(* IEC 61131-3 sources: plc-st-coding-agent/progress/evidence/f14_v10_full_20261113/jobs/codex_minimax-m27 (part 6) *)

(* ---- public-medium-08.raw_candidate_04.st ---- *)
(* ENGINEERING_CONTRACT
   PUB001: Parse dotted-decimal IPv4, validate 4 numeric segments 0-255
   PUB002: Network byte order assembly (MSB=first segment)
   PUB003: Invalid input → ipValue=0 (malformed, nondigit, wrong count, OOR)
   PUB004: Valid 0.0.0.0 also produces 0 (by assembly)

   State retention: None (stateless function block)
   Reset behavior: None (no reset input specified)
   First scan: Same as subsequent (no edge memory)

   Bug fix: Reject empty segments (consecutive delimiters like "1..2.3")
   by tracking nonempty digit accumulation per segment
*)

(* CONTRACT_RULES [] *)

FUNCTION_BLOCK IPv4_Parse
VAR_INPUT
    ipText : STRING(254);
END_VAR
VAR_OUTPUT
    ipValue : UDINT := 0;
END_VAR
VAR
    tmp_pos : UDINT;
    tmp_seg_idx : UDINT;
    tmp_char : BYTE;
    tmp_seg_val : UDINT;
    tmp_result : UDINT;
    tmp_seg_nonempty : BOOL;
END_VAR

tmp_pos := 0;
tmp_seg_idx := 0;
tmp_result := 0;
tmp_seg_val := 0;
tmp_seg_nonempty := FALSE;

WHILE tmp_pos < LEN(ipText) DO
    tmp_char := ipText[tmp_pos];

    IF tmp_char >= 48 AND tmp_char <= 57 THEN
        tmp_seg_val := tmp_seg_val * 10 + TO_UDINT(tmp_char - 48);

        IF tmp_seg_val > 255 THEN
            ipValue := 0;
            RETURN;
        END_IF;

        tmp_seg_nonempty := TRUE;
        tmp_pos := tmp_pos + 1;

    ELSIF tmp_char = 46 THEN

        IF NOT tmp_seg_nonempty THEN
            ipValue := 0;
            RETURN;
        END_IF;

        IF tmp_seg_idx >= 3 THEN
            ipValue := 0;
            RETURN;
        END_IF;

        CASE tmp_seg_idx OF
            0: tmp_result := SHL(tmp_seg_val, 24);
            1: tmp_result := tmp_result OR SHL(tmp_seg_val, 16);
            2: tmp_result := tmp_result OR SHL(tmp_seg_val, 8);
        END_CASE;

        tmp_seg_idx := tmp_seg_idx + 1;
        tmp_seg_val := 0;
        tmp_seg_nonempty := FALSE;
        tmp_pos := tmp_pos + 1;
    ELSE

        ipValue := 0;
        RETURN;
    END_IF;
END_WHILE;

IF tmp_seg_idx <> 3 THEN
    ipValue := 0;
ELSE
    tmp_result := tmp_result OR tmp_seg_val;
    ipValue := tmp_result;
END_IF;

END_FUNCTION_BLOCK

(* ---- self-easy-01.candidate_01.st ---- *)
(*
ENGINEERING_CONTRACT
================================================================
Output: avgOut (REAL)
─────────────────────────────────────────────────────────────────
Activation:    Computed every scan when enable AND avgEnable AND count > 0
Retention:     Held when enable=FALSE, avgEnable=FALSE, or count<=0
Reset:         No explicit reset; cold-start avgOut initializes to 0.0
Same-scan:     All inputs evaluated together; final timer state used
Units/bounds:  count: 0..8 clamped to 1..8 for division, sum: DINT
─────────────────────────────────────────────────────────────────
PUB001: enable=TRUE updates avgOut; enable=FALSE retains prev
PUB002: avgEnable input
PUB003: values array[1..8] of INT, 1-indexed sample storage
PUB004: count input INT
PUB005: avgOut output REAL, no rounding to integer
PUB006: count=0 -> no division by zero, avgOut unchanged
PUB007: count>8 -> use only first 8 samples, no out-of-bounds
PUB008: avgEnable=FALSE -> avgOut unchanged (retain)
PUB009: DINT/LINT summation to prevent INT overflow
PUB010: REAL output preserves original precision
================================================================
*)

(* CONTRACT_RULES [] *)

FUNCTION_BLOCK FB
VAR_INPUT
    enable    : BOOL;
    values    : ARRAY[1..8] OF INT;
    count     : INT;
    avgEnable : BOOL;
END_VAR
VAR_OUTPUT
    avgOut    : REAL := 0.0;
END_VAR
VAR
    tmp_sum   : DINT;
    tmp_count : INT;
END_VAR

tmp_count := count;
IF tmp_count < 1 THEN
    tmp_count := 0;
ELSIF tmp_count > 8 THEN
    tmp_count := 8;
END_IF;

IF enable AND avgEnable AND (tmp_count > 0) THEN
    tmp_sum := 0;
    IF tmp_count >= 1 THEN
        tmp_sum := tmp_sum + TO_DINT(values[1]);
    END_IF;
    IF tmp_count >= 2 THEN
        tmp_sum := tmp_sum + TO_DINT(values[2]);
    END_IF;
    IF tmp_count >= 3 THEN
        tmp_sum := tmp_sum + TO_DINT(values[3]);
    END_IF;
    IF tmp_count >= 4 THEN
        tmp_sum := tmp_sum + TO_DINT(values[4]);
    END_IF;
    IF tmp_count >= 5 THEN
        tmp_sum := tmp_sum + TO_DINT(values[5]);
    END_IF;
    IF tmp_count >= 6 THEN
        tmp_sum := tmp_sum + TO_DINT(values[6]);
    END_IF;
    IF tmp_count >= 7 THEN
        tmp_sum := tmp_sum + TO_DINT(values[7]);
    END_IF;
    IF tmp_count >= 8 THEN
        tmp_sum := tmp_sum + TO_DINT(values[8]);
    END_IF;
    avgOut := TO_REAL(tmp_sum) / TO_REAL(tmp_count);
END_IF;
END_FUNCTION_BLOCK

(* ---- self-easy-01.raw_candidate_01.st ---- *)
(*
ENGINEERING_CONTRACT
================================================================
Output: avgOut (REAL)
─────────────────────────────────────────────────────────────────
Activation:    Computed every scan when enable AND avgEnable AND count > 0
Retention:     Held when enable=FALSE, avgEnable=FALSE, or count<=0
Reset:         No explicit reset; cold-start avgOut initializes to 0.0
Same-scan:     All inputs evaluated together; final timer state used
Units/bounds:  count: 0..8 clamped to 1..8 for division, sum: DINT
─────────────────────────────────────────────────────────────────
PUB001: enable=TRUE updates avgOut; enable=FALSE retains prev
PUB002: avgEnable input
PUB003: values array[1..8] of INT, 1-indexed sample storage
PUB004: count input INT
PUB005: avgOut output REAL, no rounding to integer
PUB006: count=0 -> no division by zero, avgOut unchanged
PUB007: count>8 -> use only first 8 samples, no out-of-bounds
PUB008: avgEnable=FALSE -> avgOut unchanged (retain)
PUB009: DINT/LINT summation to prevent INT overflow
PUB010: REAL output preserves original precision
================================================================
*)

(* CONTRACT_RULES [] *)

FUNCTION_BLOCK FB
VAR_INPUT
    enable    : BOOL;
    values    : ARRAY[1..8] OF INT;
    count     : INT;
    avgEnable : BOOL;
END_VAR
VAR_OUTPUT
    avgOut    : REAL := 0.0;
END_VAR
VAR
    tmp_sum   : DINT;
    tmp_count : INT;
END_VAR

tmp_count := count;
IF tmp_count < 1 THEN
    tmp_count := 0;
ELSIF tmp_count > 8 THEN
    tmp_count := 8;
END_IF;

IF enable AND avgEnable AND (tmp_count > 0) THEN
    tmp_sum := 0;
    IF tmp_count >= 1 THEN
        tmp_sum := tmp_sum + TO_DINT(values[1]);
    END_IF;
    IF tmp_count >= 2 THEN
        tmp_sum := tmp_sum + TO_DINT(values[2]);
    END_IF;
    IF tmp_count >= 3 THEN
        tmp_sum := tmp_sum + TO_DINT(values[3]);
    END_IF;
    IF tmp_count >= 4 THEN
        tmp_sum := tmp_sum + TO_DINT(values[4]);
    END_IF;
    IF tmp_count >= 5 THEN
        tmp_sum := tmp_sum + TO_DINT(values[5]);
    END_IF;
    IF tmp_count >= 6 THEN
        tmp_sum := tmp_sum + TO_DINT(values[6]);
    END_IF;
    IF tmp_count >= 7 THEN
        tmp_sum := tmp_sum + TO_DINT(values[7]);
    END_IF;
    IF tmp_count >= 8 THEN
        tmp_sum := tmp_sum + TO_DINT(values[8]);
    END_IF;
    avgOut := TO_REAL(tmp_sum) / TO_REAL(tmp_count);
END_IF;
END_FUNCTION_BLOCK

(* ---- self-easy-02.candidate_01.st ---- *)
FUNCTION_BLOCK FB
VAR_INPUT
    tankLevel   : REAL;
    outletFlow  : REAL;
    inletPermit : BOOL;
    resetBtn    : BOOL;
END_VAR
VAR_OUTPUT
    pumpRun        : BOOL;
    alarmHigh      : BOOL;
    alarmLow       : BOOL;
    outletValveOpen: BOOL;
END_VAR
VAR
    prevResetBtn   : BOOL := FALSE;
    prevAlarmHigh  : BOOL := FALSE;
    prevAlarmLow   : BOOL := FALSE;
    firstScan      : BOOL := TRUE;
END_VAR
(* ENGINEERING_CONTRACT
 * ┌──────────────────┬─────────────────────────────────────────────────────────┐
 * │ alarmHigh        │ SET: tankLevel >= 85.0 (same scan priority)             │
 * │                  │ HOLD: until resetBtn rising edge AND tankLevel < 85.0   │
 * │                  │ RESET: only when safe condition cleared first           │
 * │                  │ UNITS: dimensionless % [0..100]                         │
 * ├──────────────────┼─────────────────────────────────────────────────────────┤
 * │ alarmLow         │ SET: tankLevel <= 15.0 (same scan priority)             │
 * │                  │ HOLD: until resetBtn rising edge AND tankLevel > 15.0   │
 * │                  │ RESET: only when safe condition cleared first           │
 * │                  │ UNITS: dimensionless % [0..100]                         │
 * ├──────────────────┼─────────────────────────────────────────────────────────┤
 * │ pumpRun          │ ACTIVATION: inletPermit=TRUE AND alarmHigh=FALSE AND alarmLow=FALSE │
 * │                  │ DEACTIVATION: any alarm active OR inletPermit=FALSE     │
 * │                  │ PRIORITY: stop-before-start, same-scan final state      │
 * │                  │ UNITS: command signal (BOOL)                            │
 * ├──────────────────┼─────────────────────────────────────────────────────────┤
 * │ outletValveOpen  │ ACTIVATION: alarmLow=FALSE (normal + alarmHigh-only)    │
 * │                  │ DEACTIVATION: alarmLow=TRUE                             │
 * │                  │ PRIORITY: latch follows alarmLow, no reset edge effect  │
 * │                  │ UNITS: command signal (BOOL)                            │
 * ├──────────────────┼─────────────────────────────────────────────────────────┤
 * │ resetBtn edge    │ DETECT: rising(TRUE), firstScan treated as FALSE->FALSE  │
 * │                  │ RETENTION: holding across level change does NOT trigger │
 * │                  │ UNITS: edge-detected per scan                           │
 * └──────────────────┴─────────────────────────────────────────────────────────┘
 * PUB refs: 85%/15% thresholds PUB003, latch PUB004, reset edge PUB005,
 *           pump interlock PUB006, valve PUB007, inlet permit PUB008
 *)
BEGIN
    (* Detect rising edge on resetBtn; first scan treats btn as FALSE *)
    IF firstScan THEN
        firstScan := FALSE;
    END_IF;

    (* Step 1: Update alarmHigh - immediate latch on danger condition *)
    IF tankLevel >= 85.0 THEN
        alarmHigh := TRUE;
    ELSIF resetBtn AND NOT prevResetBtn AND tankLevel < 85.0 THEN
        alarmHigh := FALSE;
    END_IF;

    (* Step 2: Update alarmLow - immediate latch on danger condition *)
    IF tankLevel <= 15.0 THEN
        alarmLow := TRUE;
    ELSIF resetBtn AND NOT prevResetBtn AND tankLevel > 15.0 THEN
        alarmLow := FALSE;
    END_IF;

    (* Step 3: pumpRun - stop before start, all conditions same scan *)
    IF alarmHigh OR alarmLow OR NOT inletPermit THEN
        pumpRun := FALSE;
    ELSE
        pumpRun := TRUE;
    END_IF;

    (* Step 4: outletValveOpen - inverse of alarmLow *)
    outletValveOpen := NOT alarmLow;

    (* Step 5: Store previous states for next scan edge detection *)
    prevResetBtn  := resetBtn;
    prevAlarmHigh := alarmHigh;
    prevAlarmLow  := alarmLow;
END_FUNCTION_BLOCK

(* ---- self-easy-02.candidate_02.st ---- *)
FUNCTION_BLOCK FB
VAR_INPUT
    tankLevel   : REAL;
    outletFlow  : REAL;
    inletPermit : BOOL;
    resetBtn    : BOOL;
END_VAR
VAR_OUTPUT
    pumpRun        : BOOL;
    alarmHigh      : BOOL;
    alarmLow       : BOOL;
    outletValveOpen: BOOL;
END_VAR
VAR
    prevResetBtn   : BOOL := FALSE;
    prevAlarmHigh  : BOOL := FALSE;
    prevAlarmLow   : BOOL := FALSE;
    firstScan      : BOOL := TRUE;
END_VAR
(* ENGINEERING_CONTRACT
 * ┌──────────────────┬─────────────────────────────────────────────────────────┐
 * │ alarmHigh        │ SET: tankLevel >= 85.0 (same scan priority)             │
 * │                  │ HOLD: until resetBtn rising edge AND tankLevel < 85.0   │
 * │                  │ RESET: only when safe condition cleared first           │
 * │                  │ UNITS: dimensionless % [0..100]                         │
 * ├──────────────────┼─────────────────────────────────────────────────────────┤
 * │ alarmLow         │ SET: tankLevel <= 15.0 (same scan priority)             │
 * │                  │ HOLD: until resetBtn rising edge AND tankLevel > 15.0   │
 * │                  │ RESET: only when safe condition cleared first           │
 * │                  │ UNITS: dimensionless % [0..100]                         │
 * ├──────────────────┼─────────────────────────────────────────────────────────┤
 * │ pumpRun          │ ACTIVATION: inletPermit=TRUE AND alarmHigh=FALSE AND alarmLow=FALSE │
 * │                  │ DEACTIVATION: any alarm active OR inletPermit=FALSE     │
 * │                  │ PRIORITY: stop-before-start, same-scan final state      │
 * │                  │ UNITS: command signal (BOOL)                            │
 * ├──────────────────┼─────────────────────────────────────────────────────────┤
 * │ outletValveOpen  │ ACTIVATION: alarmLow=FALSE (normal + alarmHigh-only)    │
 * │                  │ DEACTIVATION: alarmLow=TRUE                             │
 * │                  │ PRIORITY: latch follows alarmLow, no reset edge effect  │
 * │                  │ UNITS: command signal (BOOL)                            │
 * ├──────────────────┼─────────────────────────────────────────────────────────┤
 * │ resetBtn edge    │ DETECT: rising(TRUE), firstScan treated as FALSE->FALSE  │
 * │                  │ RETENTION: holding across level change does NOT trigger │
 * │                  │ UNITS: edge-detected per scan                           │
 * └──────────────────┴─────────────────────────────────────────────────────────┘
 * PUB refs: 85%/15% thresholds PUB003, latch PUB004, reset edge PUB005,
 *           pump interlock PUB006, valve PUB007, inlet permit PUB008
 *)
BEGIN
    (* Step 1: Update alarmHigh - immediate latch on danger condition *)
    IF tankLevel >= 85.0 THEN
        alarmHigh := TRUE;
    ELSIF resetBtn AND NOT prevResetBtn AND NOT firstScan AND tankLevel < 85.0 THEN
        alarmHigh := FALSE;
    END_IF;

    (* Step 2: Update alarmLow - immediate latch on danger condition *)
    IF tankLevel <= 15.0 THEN
        alarmLow := TRUE;
    ELSIF resetBtn AND NOT prevResetBtn AND NOT firstScan AND tankLevel > 15.0 THEN
        alarmLow := FALSE;
    END_IF;

    (* Step 3: pumpRun - stop before start, all conditions same scan *)
    IF alarmHigh OR alarmLow OR NOT inletPermit THEN
        pumpRun := FALSE;
    ELSE
        pumpRun := TRUE;
    END_IF;

    (* Step 4: outletValveOpen - inverse of alarmLow *)
    outletValveOpen := NOT alarmLow;

    (* Step 5: Store previous states for next scan *)
    prevResetBtn  := resetBtn;
    prevAlarmHigh := alarmHigh;
    prevAlarmLow  := alarmLow;
    firstScan     := FALSE;
END_FUNCTION_BLOCK

(* ---- self-easy-02.candidate_03.st ---- *)
FUNCTION_BLOCK FB
VAR_INPUT
    tankLevel   : REAL;
    outletFlow  : REAL;
    inletPermit : BOOL;
    resetBtn    : BOOL;
END_VAR
VAR_OUTPUT
    pumpRun        : BOOL;
    alarmHigh      : BOOL;
    alarmLow       : BOOL;
    outletValveOpen: BOOL;
END_VAR
VAR
    prevResetBtn : BOOL := FALSE;
END_VAR
(* ENGINEERING_CONTRACT *)
(* alarmHigh: SET at tankLevel>=85.0 (same-scan priority). HOLD until resetBtn rising AND tankLevel<85.0. RESET only when safe first. *)
(* alarmLow:  SET at tankLevel<=15.0 (same-scan priority). HOLD until resetBtn rising AND tankLevel>15.0. RESET only when safe first. *)
(* pumpRun:   ACT when inletPermit=TRUE AND alarmHigh=FALSE AND alarmLow=FALSE. STOP on any alarm or !inletPermit. *)
(* outletValveOpen: ON when alarmLow=FALSE. OFF when alarmLow=TRUE. No reset edge effect. *)
(* resetBtn:  Rising edge detection, firstScan=FALSE. Holding across level change does NOT re-trigger. *)
BEGIN
    (* Update alarmHigh *)
    IF tankLevel >= 85.0 THEN
        alarmHigh := TRUE;
    ELSIF resetBtn AND NOT prevResetBtn AND tankLevel < 85.0 THEN
        alarmHigh := FALSE;
    END_IF;

    (* Update alarmLow *)
    IF tankLevel <= 15.0 THEN
        alarmLow := TRUE;
    ELSIF resetBtn AND NOT prevResetBtn AND tankLevel > 15.0 THEN
        alarmLow := FALSE;
    END_IF;

    (* pumpRun: stop before start *)
    IF alarmHigh OR alarmLow OR NOT inletPermit THEN
        pumpRun := FALSE;
    ELSE
        pumpRun := TRUE;
    END_IF;

    (* outletValveOpen: inverse of alarmLow *)
    outletValveOpen := NOT alarmLow;

    (* Store previous state *)
    prevResetBtn := resetBtn;
END_FUNCTION_BLOCK
(* CONTRACT_RULES [] *)

(* ---- self-easy-02.candidate_04.st ---- *)
FUNCTION_BLOCK FB
VAR_INPUT
    tankLevel   : REAL;
    outletFlow  : REAL;
    inletPermit : BOOL;
    resetBtn    : BOOL;
END_VAR
VAR_OUTPUT
    pumpRun        : BOOL;
    alarmHigh      : BOOL;
    alarmLow       : BOOL;
    outletValveOpen: BOOL;
END_VAR
VAR
    prevResetBtn   : BOOL := FALSE;
    firstScan      : BOOL := TRUE;
END_VAR
(* ENGINEERING_CONTRACT
 * ┌──────────────────┬─────────────────────────────────────────────────────────┐
 * │ alarmHigh        │ SET: tankLevel >= 85.0 (same scan priority)             │
 * │                  │ HOLD: until resetBtn rising edge AND tankLevel < 85.0   │
 * │                  │ RESET: only when safe condition cleared first           │
 * │                  │ UNITS: dimensionless % [0..100]                         │
 * ├──────────────────┼─────────────────────────────────────────────────────────┤
 * │ alarmLow         │ SET: tankLevel <= 15.0 (same scan priority)             │
 * │                  │ HOLD: until resetBtn rising edge AND tankLevel > 15.0   │
 * │                  │ RESET: only when safe condition cleared first           │
 * │                  │ UNITS: dimensionless % [0..100]                         │
 * ├──────────────────┼─────────────────────────────────────────────────────────┤
 * │ pumpRun          │ ACTIVATION: inletPermit=TRUE AND alarmHigh=FALSE AND alarmLow=FALSE │
 * │                  │ DEACTIVATION: any alarm active OR inletPermit=FALSE     │
 * │                  │ PRIORITY: stop-before-start, same-scan final state      │
 * │                  │ UNITS: command signal (BOOL)                            │
 * ├──────────────────┼─────────────────────────────────────────────────────────┤
 * │ outletValveOpen  │ ACTIVATION: alarmLow=FALSE (normal + alarmHigh-only)    │
 * │                  │ DEACTIVATION: alarmLow=TRUE                             │
 * │                  │ PRIORITY: latch follows alarmLow, no reset edge effect  │
 * │                  │ UNITS: command signal (BOOL)                            │
 * ├──────────────────┼─────────────────────────────────────────────────────────┤
 * │ resetBtn edge    │ DETECT: rising(TRUE), firstScan treated as FALSE->FALSE  │
 * │                  │ RETENTION: holding across level change does NOT trigger │
 * │                  │ UNITS: edge-detected per scan                           │
 * └──────────────────┴─────────────────────────────────────────────────────────┘
 * PUB refs: 85%/15% thresholds PUB003, latch PUB004, reset edge PUB005,
 *           pump interlock PUB006, valve PUB007, inlet permit PUB008
 *)
BEGIN
    IF firstScan THEN
        firstScan := FALSE;
        prevResetBtn := FALSE;
    END_IF;

    IF tankLevel >= 85.0 THEN
        alarmHigh := TRUE;
    ELSIF resetBtn AND NOT prevResetBtn AND tankLevel < 85.0 THEN
        alarmHigh := FALSE;
    END_IF;

    IF tankLevel <= 15.0 THEN
        alarmLow := TRUE;
    ELSIF resetBtn AND NOT prevResetBtn AND tankLevel > 15.0 THEN
        alarmLow := FALSE;
    END_IF;

    IF alarmHigh OR alarmLow OR NOT inletPermit THEN
        pumpRun := FALSE;
    ELSE
        pumpRun := TRUE;
    END_IF;

    outletValveOpen := NOT alarmLow;

    prevResetBtn := resetBtn;
END_FUNCTION_BLOCK
(* CONTRACT_RULES [] *)

(* ---- self-easy-02.raw_candidate_01.st ---- *)
FUNCTION_BLOCK FB
VAR_INPUT
    tankLevel   : REAL;
    outletFlow  : REAL;
    inletPermit : BOOL;
    resetBtn    : BOOL;
END_VAR
VAR_OUTPUT
    pumpRun        : BOOL;
    alarmHigh      : BOOL;
    alarmLow       : BOOL;
    outletValveOpen: BOOL;
END_VAR
VAR
    prevResetBtn   : BOOL := FALSE;
    prevAlarmHigh  : BOOL := FALSE;
    prevAlarmLow   : BOOL := FALSE;
    firstScan      : BOOL := TRUE;
END_VAR
(* ENGINEERING_CONTRACT
 * ┌──────────────────┬─────────────────────────────────────────────────────────┐
 * │ alarmHigh        │ SET: tankLevel >= 85.0 (same scan priority)             │
 * │                  │ HOLD: until resetBtn rising edge AND tankLevel < 85.0   │
 * │                  │ RESET: only when safe condition cleared first           │
 * │                  │ UNITS: dimensionless % [0..100]                         │
 * ├──────────────────┼─────────────────────────────────────────────────────────┤
 * │ alarmLow         │ SET: tankLevel <= 15.0 (same scan priority)             │
 * │                  │ HOLD: until resetBtn rising edge AND tankLevel > 15.0   │
 * │                  │ RESET: only when safe condition cleared first           │
 * │                  │ UNITS: dimensionless % [0..100]                         │
 * ├──────────────────┼─────────────────────────────────────────────────────────┤
 * │ pumpRun          │ ACTIVATION: inletPermit=TRUE AND alarmHigh=FALSE AND alarmLow=FALSE │
 * │                  │ DEACTIVATION: any alarm active OR inletPermit=FALSE     │
 * │                  │ PRIORITY: stop-before-start, same-scan final state      │
 * │                  │ UNITS: command signal (BOOL)                            │
 * ├──────────────────┼─────────────────────────────────────────────────────────┤
 * │ outletValveOpen  │ ACTIVATION: alarmLow=FALSE (normal + alarmHigh-only)    │
 * │                  │ DEACTIVATION: alarmLow=TRUE                             │
 * │                  │ PRIORITY: latch follows alarmLow, no reset edge effect  │
 * │                  │ UNITS: command signal (BOOL)                            │
 * ├──────────────────┼─────────────────────────────────────────────────────────┤
 * │ resetBtn edge    │ DETECT: rising(TRUE), firstScan treated as FALSE->FALSE  │
 * │                  │ RETENTION: holding across level change does NOT trigger │
 * │                  │ UNITS: edge-detected per scan                           │
 * └──────────────────┴─────────────────────────────────────────────────────────┘
 * PUB refs: 85%/15% thresholds PUB003, latch PUB004, reset edge PUB005,
 *           pump interlock PUB006, valve PUB007, inlet permit PUB008
 *)
BEGIN
    (* Detect rising edge on resetBtn; first scan treats btn as FALSE *)
    IF firstScan THEN
        firstScan := FALSE;
    END_IF;

    (* Step 1: Update alarmHigh - immediate latch on danger condition *)
    IF tankLevel >= 85.0 THEN
        alarmHigh := TRUE;
    ELSIF resetBtn AND NOT prevResetBtn AND tankLevel < 85.0 THEN
        alarmHigh := FALSE;
    END_IF;

    (* Step 2: Update alarmLow - immediate latch on danger condition *)
    IF tankLevel <= 15.0 THEN
        alarmLow := TRUE;
    ELSIF resetBtn AND NOT prevResetBtn AND tankLevel > 15.0 THEN
        alarmLow := FALSE;
    END_IF;

    (* Step 3: pumpRun - stop before start, all conditions same scan *)
    IF alarmHigh OR alarmLow OR NOT inletPermit THEN
        pumpRun := FALSE;
    ELSE
        pumpRun := TRUE;
    END_IF;

    (* Step 4: outletValveOpen - inverse of alarmLow *)
    outletValveOpen := NOT alarmLow;

    (* Step 5: Store previous states for next scan edge detection *)
    prevResetBtn  := resetBtn;
    prevAlarmHigh := alarmHigh;
    prevAlarmLow  := alarmLow;
END_FUNCTION_BLOCK

(* ---- self-easy-02.raw_candidate_02.st ---- *)
FUNCTION_BLOCK FB
VAR_INPUT
    tankLevel   : REAL;
    outletFlow  : REAL;
    inletPermit : BOOL;
    resetBtn    : BOOL;
END_VAR
VAR_OUTPUT
    pumpRun        : BOOL;
    alarmHigh      : BOOL;
    alarmLow       : BOOL;
    outletValveOpen: BOOL;
END_VAR
VAR
    prevResetBtn   : BOOL := FALSE;
    prevAlarmHigh  : BOOL := FALSE;
    prevAlarmLow   : BOOL := FALSE;
    firstScan      : BOOL := TRUE;
END_VAR
(* ENGINEERING_CONTRACT
 * ┌──────────────────┬─────────────────────────────────────────────────────────┐
 * │ alarmHigh        │ SET: tankLevel >= 85.0 (same scan priority)             │
 * │                  │ HOLD: until resetBtn rising edge AND tankLevel < 85.0   │
 * │                  │ RESET: only when safe condition cleared first           │
 * │                  │ UNITS: dimensionless % [0..100]                         │
 * ├──────────────────┼─────────────────────────────────────────────────────────┤
 * │ alarmLow         │ SET: tankLevel <= 15.0 (same scan priority)             │
 * │                  │ HOLD: until resetBtn rising edge AND tankLevel > 15.0   │
 * │                  │ RESET: only when safe condition cleared first           │
 * │                  │ UNITS: dimensionless % [0..100]                         │
 * ├──────────────────┼─────────────────────────────────────────────────────────┤
 * │ pumpRun          │ ACTIVATION: inletPermit=TRUE AND alarmHigh=FALSE AND alarmLow=FALSE │
 * │                  │ DEACTIVATION: any alarm active OR inletPermit=FALSE     │
 * │                  │ PRIORITY: stop-before-start, same-scan final state      │
 * │                  │ UNITS: command signal (BOOL)                            │
 * ├──────────────────┼─────────────────────────────────────────────────────────┤
 * │ outletValveOpen  │ ACTIVATION: alarmLow=FALSE (normal + alarmHigh-only)    │
 * │                  │ DEACTIVATION: alarmLow=TRUE                             │
 * │                  │ PRIORITY: latch follows alarmLow, no reset edge effect  │
 * │                  │ UNITS: command signal (BOOL)                            │
 * ├──────────────────┼─────────────────────────────────────────────────────────┤
 * │ resetBtn edge    │ DETECT: rising(TRUE), firstScan treated as FALSE->FALSE  │
 * │                  │ RETENTION: holding across level change does NOT trigger │
 * │                  │ UNITS: edge-detected per scan                           │
 * └──────────────────┴─────────────────────────────────────────────────────────┘
 * PUB refs: 85%/15% thresholds PUB003, latch PUB004, reset edge PUB005,
 *           pump interlock PUB006, valve PUB007, inlet permit PUB008
 *)
BEGIN
    (* Step 1: Update alarmHigh - immediate latch on danger condition *)
    IF tankLevel >= 85.0 THEN
        alarmHigh := TRUE;
    ELSIF resetBtn AND NOT prevResetBtn AND NOT firstScan AND tankLevel < 85.0 THEN
        alarmHigh := FALSE;
    END_IF;

    (* Step 2: Update alarmLow - immediate latch on danger condition *)
    IF tankLevel <= 15.0 THEN
        alarmLow := TRUE;
    ELSIF resetBtn AND NOT prevResetBtn AND NOT firstScan AND tankLevel > 15.0 THEN
        alarmLow := FALSE;
    END_IF;

    (* Step 3: pumpRun - stop before start, all conditions same scan *)
    IF alarmHigh OR alarmLow OR NOT inletPermit THEN
        pumpRun := FALSE;
    ELSE
        pumpRun := TRUE;
    END_IF;

    (* Step 4: outletValveOpen - inverse of alarmLow *)
    outletValveOpen := NOT alarmLow;

    (* Step 5: Store previous states for next scan *)
    prevResetBtn  := resetBtn;
    prevAlarmHigh := alarmHigh;
    prevAlarmLow  := alarmLow;
    firstScan     := FALSE;
END_FUNCTION_BLOCK

(* ---- self-easy-02.raw_candidate_03.st ---- *)
FUNCTION_BLOCK FB
VAR_INPUT
    tankLevel   : REAL;
    outletFlow  : REAL;
    inletPermit : BOOL;
    resetBtn    : BOOL;
END_VAR
VAR_OUTPUT
    pumpRun        : BOOL;
    alarmHigh      : BOOL;
    alarmLow       : BOOL;
    outletValveOpen: BOOL;
END_VAR
VAR
    prevResetBtn : BOOL := FALSE;
END_VAR
(* ENGINEERING_CONTRACT *)
(* alarmHigh: SET at tankLevel>=85.0 (same-scan priority). HOLD until resetBtn rising AND tankLevel<85.0. RESET only when safe first. *)
(* alarmLow:  SET at tankLevel<=15.0 (same-scan priority). HOLD until resetBtn rising AND tankLevel>15.0. RESET only when safe first. *)
(* pumpRun:   ACT when inletPermit=TRUE AND alarmHigh=FALSE AND alarmLow=FALSE. STOP on any alarm or !inletPermit. *)
(* outletValveOpen: ON when alarmLow=FALSE. OFF when alarmLow=TRUE. No reset edge effect. *)
(* resetBtn:  Rising edge detection, firstScan=FALSE. Holding across level change does NOT re-trigger. *)
BEGIN
    (* Update alarmHigh *)
    IF tankLevel >= 85.0 THEN
        alarmHigh := TRUE;
    ELSIF resetBtn AND NOT prevResetBtn AND tankLevel < 85.0 THEN
        alarmHigh := FALSE;
    END_IF;

    (* Update alarmLow *)
    IF tankLevel <= 15.0 THEN
        alarmLow := TRUE;
    ELSIF resetBtn AND NOT prevResetBtn AND tankLevel > 15.0 THEN
        alarmLow := FALSE;
    END_IF;

    (* pumpRun: stop before start *)
    IF alarmHigh OR alarmLow OR NOT inletPermit THEN
        pumpRun := FALSE;
    ELSE
        pumpRun := TRUE;
    END_IF;

    (* outletValveOpen: inverse of alarmLow *)
    outletValveOpen := NOT alarmLow;

    (* Store previous state *)
    prevResetBtn := resetBtn;
END_FUNCTION_BLOCK
(* CONTRACT_RULES [] *)

(* ---- self-easy-02.raw_candidate_04.st ---- *)
FUNCTION_BLOCK FB
VAR_INPUT
    tankLevel   : REAL;
    outletFlow  : REAL;
    inletPermit : BOOL;
    resetBtn    : BOOL;
END_VAR
VAR_OUTPUT
    pumpRun        : BOOL;
    alarmHigh      : BOOL;
    alarmLow       : BOOL;
    outletValveOpen: BOOL;
END_VAR
VAR
    prevResetBtn   : BOOL := FALSE;
    firstScan      : BOOL := TRUE;
END_VAR
(* ENGINEERING_CONTRACT
 * ┌──────────────────┬─────────────────────────────────────────────────────────┐
 * │ alarmHigh        │ SET: tankLevel >= 85.0 (same scan priority)             │
 * │                  │ HOLD: until resetBtn rising edge AND tankLevel < 85.0   │
 * │                  │ RESET: only when safe condition cleared first           │
 * │                  │ UNITS: dimensionless % [0..100]                         │
 * ├──────────────────┼─────────────────────────────────────────────────────────┤
 * │ alarmLow         │ SET: tankLevel <= 15.0 (same scan priority)             │
 * │                  │ HOLD: until resetBtn rising edge AND tankLevel > 15.0   │
 * │                  │ RESET: only when safe condition cleared first           │
 * │                  │ UNITS: dimensionless % [0..100]                         │
 * ├──────────────────┼─────────────────────────────────────────────────────────┤
 * │ pumpRun          │ ACTIVATION: inletPermit=TRUE AND alarmHigh=FALSE AND alarmLow=FALSE │
 * │                  │ DEACTIVATION: any alarm active OR inletPermit=FALSE     │
 * │                  │ PRIORITY: stop-before-start, same-scan final state      │
 * │                  │ UNITS: command signal (BOOL)                            │
 * ├──────────────────┼─────────────────────────────────────────────────────────┤
 * │ outletValveOpen  │ ACTIVATION: alarmLow=FALSE (normal + alarmHigh-only)    │
 * │                  │ DEACTIVATION: alarmLow=TRUE                             │
 * │                  │ PRIORITY: latch follows alarmLow, no reset edge effect  │
 * │                  │ UNITS: command signal (BOOL)                            │
 * ├──────────────────┼─────────────────────────────────────────────────────────┤
 * │ resetBtn edge    │ DETECT: rising(TRUE), firstScan treated as FALSE->FALSE  │
 * │                  │ RETENTION: holding across level change does NOT trigger │
 * │                  │ UNITS: edge-detected per scan                           │
 * └──────────────────┴─────────────────────────────────────────────────────────┘
 * PUB refs: 85%/15% thresholds PUB003, latch PUB004, reset edge PUB005,
 *           pump interlock PUB006, valve PUB007, inlet permit PUB008
 *)
BEGIN
    IF firstScan THEN
        firstScan := FALSE;
        prevResetBtn := FALSE;
    END_IF;

    IF tankLevel >= 85.0 THEN
        alarmHigh := TRUE;
    ELSIF resetBtn AND NOT prevResetBtn AND tankLevel < 85.0 THEN
        alarmHigh := FALSE;
    END_IF;

    IF tankLevel <= 15.0 THEN
        alarmLow := TRUE;
    ELSIF resetBtn AND NOT prevResetBtn AND tankLevel > 15.0 THEN
        alarmLow := FALSE;
    END_IF;

    IF alarmHigh OR alarmLow OR NOT inletPermit THEN
        pumpRun := FALSE;
    ELSE
        pumpRun := TRUE;
    END_IF;

    outletValveOpen := NOT alarmLow;

    prevResetBtn := resetBtn;
END_FUNCTION_BLOCK
(* CONTRACT_RULES [] *)

(* ---- self-hard-01.candidate_01.st ---- *)
FUNCTION_BLOCK FB
VAR_INPUT
    flowLow   : BOOL;
    ackBtn    : BOOL;
    sensorOK  : BOOL;
END_VAR
VAR_OUTPUT
    alarmActive : BOOL;
    alarmAcked  : BOOL;
    highHigh    : BOOL;
END_VAR
VAR
    prev_flowLow : BOOL := FALSE;
    prev_ackBtn  : BOOL := FALSE;
    tmp_flowRising : BOOL;
    tmp_ackRising  : BOOL;
END_VAR

(*
ENGINEERING_CONTRACT:
================================================================================
| Output/State        | Activation          | Retention      | Reset/Deact         | Scan Priority | Units/Range       |
|---------------------|---------------------|----------------|---------------------|---------------|-------------------|
| alarmActive [BOOL]  | flowLow rising edge | Until explicit | rising(ackBtn) + !flowLow + tmp_unacked_wait; | Same-scan | 0..1 |
|                     |                     | deactivation   | tmp_unacked_wait := TRUE on flowLow falling  |               |                   |
|                     |                     |                | while !alarmAcked                         |               |                   |
| alarmAcked [BOOL]   | rising(ackBtn) with | Cleared on new | rising(ackBtn) + !flowLow + tmp_unacked_wait | Same-scan | 0..1 |
|                     | flowLow present;    | flowLow rise;  |                                             |               |                   |
|                     | flowLow fall while  | retained during|                                             |               |                   |
|                     | !alarmAcked         | waiting state  |                                             |               |                   |
| highHigh [BOOL]     | !sensorOK (PUB027)  | Retained while | sensorOK TRUE (PUB035)                     | Same-scan | 0..1 |
|                     |                     | !sensorOK      |                                             |               |                   |
| tmp_unacked_wait    | flowLow falling     | Until rising   | rising(ackBtn) + !flowLow                  | Internal  | Named boolean     |
| [BOOL, local]       | while !alarmAcked   | (ackBtn)       |                                             |           |                   |
================================================================================
PUB IDs: alarmActive→PUB001/PUB002/PUB003/PUB004/PUB005/PUB006; alarmAcked→PUB007/PUB008/PUB009/PUB010/PUB011/PUB012; highHigh→PUB027/PUB035

CONTRACT_RULES: []
================================================================================
*)

tmp_flowRising := flowLow AND NOT prev_flowLow;
tmp_ackRising  := ackBtn  AND NOT prev_ackBtn;

alarmActive := alarmActive;
alarmAcked  := alarmAcked;

IF tmp_flowRising THEN
    alarmActive := TRUE;
    alarmAcked  := FALSE;
ELSIF alarmActive AND tmp_ackRising THEN
    IF NOT flowLow THEN
        alarmActive := FALSE;
        alarmAcked  := FALSE;
    ELSE
        alarmAcked  := TRUE;
    END_IF;
ELSIF alarmActive AND NOT flowLow AND NOT alarmAcked THEN
    alarmAcked := TRUE;
ELSIF alarmActive AND flowLow AND alarmAcked AND tmp_flowRising THEN
    alarmAcked := FALSE;
END_IF;

highHigh := NOT sensorOK;

prev_flowLow := flowLow;
prev_ackBtn  := ackBtn;

END_FUNCTION_BLOCK

(* ---- self-hard-01.candidate_02.st ---- *)
FUNCTION_BLOCK FB
VAR_INPUT
    flowLow   : BOOL;
    ackBtn    : BOOL;
    sensorOK  : BOOL;
END_VAR
VAR_OUTPUT
    alarmActive : BOOL;
    alarmAcked  : BOOL;
    highHigh    : BOOL;
END_VAR
VAR
    prev_flowLow : BOOL := FALSE;
    tmp_flowRising : BOOL;
    tmp_ackRising  : BOOL;
END_VAR

(*
ENGINEERING_CONTRACT:
================================================================================
| Output/State        | Activation          | Retention      | Reset/Deact         | Scan Priority | Units/Range       |
|---------------------|---------------------|----------------|---------------------|---------------|-------------------|
| alarmActive [BOOL]  | flowLow rising edge | Until explicit | rising(ackBtn)+!flowLow+tmp_unacked_wait| Same-scan | 0..1 |
|                     |                     | deactivation   | tmp_unacked_wait:=TRUE on flowLow fall  |               |                   |
|                     |                     |                | while !alarmAcked                         |               |                   |
| alarmAcked [BOOL]   | rising(ackBtn) with | Cleared on new | rising(ackBtn)+!flowLow+tmp_unacked_wait | Same-scan | 0..1 |
|                     | flowLow present;    | flowLow rise;  |                                             |               |                   |
|                     | flowLow fall while  | retained during|                                             |               |                   |
|                     | !alarmAcked         | waiting state  |                                             |               |                   |
| highHigh [BOOL]     | !sensorOK (PUB027)  | Retained while | sensorOK TRUE (PUB035)                     | Same-scan | 0..1 |
|                     |                     | !sensorOK      |                                             |               |                   |
| tmp_unacked_wait    | flowLow falling     | Until rising   | rising(ackBtn)+!flowLow                  | Internal  | Named boolean     |
| [BOOL, local]       | while !alarmAcked   | (ackBtn)       |                                             |           |                   |
================================================================================
PUB IDs: alarmActive→PUB001/PUB002/PUB003/PUB004/PUB005/PUB006; alarmAcked→PUB007/PUB008/PUB009/PUB010/PUB011/PUB012; highHigh→PUB027/PUB035

CONTRACT_RULES: []
================================================================================
*)

tmp_flowRising := flowLow AND NOT prev_flowLow;
tmp_ackRising  := ackBtn  AND NOT prev_ackBtn;

IF tmp_flowRising THEN
    alarmActive := TRUE;
    alarmAcked  := FALSE;
ELSIF alarmActive AND tmp_ackRising THEN
    IF NOT flowLow THEN
        alarmActive := FALSE;
        alarmAcked  := FALSE;
    ELSE
        alarmAcked  := TRUE;
    END_IF;
ELSIF alarmActive AND NOT flowLow AND NOT alarmAcked AND prev_flowLow THEN
    alarmAcked := TRUE;
ELSIF alarmActive AND flowLow AND alarmAcked AND tmp_flowRising THEN
    alarmAcked := FALSE;
END_IF;

highHigh := NOT sensorOK;

prev_flowLow := flowLow;
prev_ackBtn  := ackBtn;

END_FUNCTION_BLOCK

(* ---- self-hard-01.candidate_03.st ---- *)
FUNCTION_BLOCK FB
VAR_INPUT
    flowLow   : BOOL;
    ackBtn    : BOOL;
    sensorOK  : BOOL;
END_VAR
VAR_OUTPUT
    alarmActive : BOOL;
    alarmAcked  : BOOL;
    highHigh    : BOOL;
END_VAR
VAR
    prev_flowLow : BOOL := FALSE;
    prev_ackBtn  : BOOL := FALSE;
    tmp_flowRising : BOOL;
    tmp_ackRising  : BOOL;
END_VAR

(*
ENGINEERING_CONTRACT:
================================================================================
| Output/State        | Activation          | Retention      | Reset/Deact         | Scan Priority | Units/Range       |
|---------------------|---------------------|----------------|---------------------|---------------|-------------------|
| alarmActive [BOOL]  | flowLow rising edge | Until explicit | rising(ackBtn)+!flowLow; or flowLow | Same-scan | 0..1 |
|                     | (PUB001)            | deactivation   | rises while alarmAcked=TRUE (new occ) |          |                   |
| alarmAcked [BOOL]   | rising(ackBtn) with | Cleared on new | rising(ackBtn)+!flowLow (PUB009/PUB010) | Same-scan | 0..1 |
|                     | flowLow present     | flowLow rise   |                                         |               |                   |
|                     | (PUB008/PUB011);    | (new occ)      |                                         |               |                   |
|                     | flowLow falling     | Retained while |                                         |               |                   |
|                     | while !alarmAcked   | waiting clear  |                                         |               |                   |
|                     | (PUB006: pending)   | (PUB006)       |                                         |               |                   |
| highHigh [BOOL]     | !sensorOK (PUB027)  | Retained while | sensorOK TRUE (PUB035)                  | Same-scan | 0..1 |
|                     |                     | !sensorOK      |                                         |               |                   |
================================================================================
PUB IDs: alarmActive→PUB001/PUB002/PUB003/PUB004/PUB005/PUB006;
         alarmAcked→PUB006/PUB007/PUB008/PUB009/PUB010/PUB011/PUB012;
         highHigh→PUB027/PUB035

CONTRACT_RULES: []
================================================================================
*)

tmp_flowRising := flowLow AND NOT prev_flowLow;
tmp_ackRising  := ackBtn  AND NOT prev_ackBtn;

IF tmp_flowRising THEN
    alarmActive := TRUE;
    alarmAcked  := FALSE;
ELSIF alarmActive AND tmp_ackRising THEN
    IF NOT flowLow THEN
        alarmActive := FALSE;
        alarmAcked  := FALSE;
    ELSE
        alarmAcked  := TRUE;
    END_IF;
ELSIF alarmActive AND NOT flowLow AND NOT alarmAcked THEN
    alarmAcked := TRUE;
ELSIF alarmActive AND NOT flowLow AND alarmAcked THEN
    alarmActive := FALSE;
    alarmAcked  := FALSE;
END_IF;

highHigh := NOT sensorOK;

prev_flowLow := flowLow;
prev_ackBtn  := ackBtn;

END_FUNCTION_BLOCK

(* ---- self-hard-01.candidate_04.st ---- *)
FUNCTION_BLOCK FB
VAR_INPUT
    flowLow   : BOOL;
    ackBtn    : BOOL;
    sensorOK  : BOOL;
END_VAR
VAR_OUTPUT
    alarmActive : BOOL;
    alarmAcked  : BOOL;
    highHigh    : BOOL;
END_VAR
VAR
    prev_flowLow : BOOL := FALSE;
    prev_ackBtn  : BOOL := FALSE;
    tmp_flowRising : BOOL;
    tmp_ackRising  : BOOL;
END_VAR

(*
ENGINEERING_CONTRACT:
================================================================================
| Output/State        | Activation          | Retention      | Reset/Deact         | Scan Priority | Units/Range       |
|---------------------|---------------------|----------------|---------------------|---------------|-------------------|
| alarmActive [BOOL]  | flowLow rising edge | Until explicit | rising(ackBtn)+!flowLow; or flowLow | Same-scan | 0..1 |
|                     | (PUB001)            | deactivation   | rises while alarmAcked=TRUE (new occ) |          |                   |
| alarmAcked [BOOL]   | rising(ackBtn) with | Cleared on new | rising(ackBtn)+!flowLow (PUB009/PUB010) | Same-scan | 0..1 |
|                     | flowLow present     | flowLow rise   |                                         |               |                   |
|                     | (PUB008/PUB011);    | (new occ)      |                                         |               |                   |
|                     | flowLow falling     | Retained while |                                         |               |                   |
|                     | while !alarmAcked   | waiting clear  |                                         |               |                   |
|                     | (PUB006: pending)   | (PUB006)       |                                         |               |                   |
| highHigh [BOOL]     | !sensorOK (PUB027)  | Retained while | sensorOK TRUE (PUB035)                  | Same-scan | 0..1 |
|                     |                     | !sensorOK      |                                         |               |                   |
================================================================================
PUB IDs: alarmActive→PUB001/PUB002/PUB003/PUB004/PUB005/PUB006;
         alarmAcked→PUB006/PUB007/PUB008/PUB009/PUB010/PUB011/PUB012;
         highHigh→PUB027/PUB035

CONTRACT_RULES: []
================================================================================
*)

tmp_flowRising := flowLow AND NOT prev_flowLow;
tmp_ackRising  := ackBtn  AND NOT prev_ackBtn;

IF tmp_flowRising THEN
    alarmActive := TRUE;
    alarmAcked  := FALSE;
ELSIF alarmActive AND tmp_ackRising AND (flowLow OR alarmAcked) THEN
    alarmAcked := TRUE;
ELSIF alarmActive AND NOT flowLow AND NOT alarmAcked THEN
    alarmAcked := TRUE;
ELSIF alarmActive AND NOT flowLow THEN
    alarmActive := FALSE;
    alarmAcked  := FALSE;
END_IF;

highHigh := NOT sensorOK;

prev_flowLow := flowLow;
prev_ackBtn  := ackBtn;

END_FUNCTION_BLOCK

(* ---- self-hard-01.raw_candidate_01.st ---- *)
FUNCTION_BLOCK FB
VAR_INPUT
    flowLow   : BOOL;
    ackBtn    : BOOL;
    sensorOK  : BOOL;
END_VAR
VAR_OUTPUT
    alarmActive : BOOL;
    alarmAcked  : BOOL;
    highHigh    : BOOL;
END_VAR
VAR
    prev_flowLow : BOOL := FALSE;
    prev_ackBtn  : BOOL := FALSE;
    tmp_flowRising : BOOL;
    tmp_ackRising  : BOOL;
END_VAR

(*
ENGINEERING_CONTRACT:
================================================================================
| Output/State        | Activation          | Retention      | Reset/Deact         | Scan Priority | Units/Range       |
|---------------------|---------------------|----------------|---------------------|---------------|-------------------|
| alarmActive [BOOL]  | flowLow rising edge | Until explicit | rising(ackBtn) + !flowLow + tmp_unacked_wait; | Same-scan | 0..1 |
|                     |                     | deactivation   | tmp_unacked_wait := TRUE on flowLow falling  |               |                   |
|                     |                     |                | while !alarmAcked                         |               |                   |
| alarmAcked [BOOL]   | rising(ackBtn) with | Cleared on new | rising(ackBtn) + !flowLow + tmp_unacked_wait | Same-scan | 0..1 |
|                     | flowLow present;    | flowLow rise;  |                                             |               |                   |
|                     | flowLow fall while  | retained during|                                             |               |                   |
|                     | !alarmAcked         | waiting state  |                                             |               |                   |
| highHigh [BOOL]     | !sensorOK (PUB027)  | Retained while | sensorOK TRUE (PUB035)                     | Same-scan | 0..1 |
|                     |                     | !sensorOK      |                                             |               |                   |
| tmp_unacked_wait    | flowLow falling     | Until rising   | rising(ackBtn) + !flowLow                  | Internal  | Named boolean     |
| [BOOL, local]       | while !alarmAcked   | (ackBtn)       |                                             |           |                   |
================================================================================
PUB IDs: alarmActive→PUB001/PUB002/PUB003/PUB004/PUB005/PUB006; alarmAcked→PUB007/PUB008/PUB009/PUB010/PUB011/PUB012; highHigh→PUB027/PUB035

CONTRACT_RULES: []
================================================================================
*)

tmp_flowRising := flowLow AND NOT prev_flowLow;
tmp_ackRising  := ackBtn  AND NOT prev_ackBtn;

alarmActive := alarmActive;
alarmAcked  := alarmAcked;

IF tmp_flowRising THEN
    alarmActive := TRUE;
    alarmAcked  := FALSE;
ELSIF alarmActive AND tmp_ackRising THEN
    IF NOT flowLow THEN
        alarmActive := FALSE;
        alarmAcked  := FALSE;
    ELSE
        alarmAcked  := TRUE;
    END_IF;
ELSIF alarmActive AND NOT flowLow AND NOT alarmAcked THEN
    alarmAcked := TRUE;
ELSIF alarmActive AND flowLow AND alarmAcked AND tmp_flowRising THEN
    alarmAcked := FALSE;
END_IF;

highHigh := NOT sensorOK;

prev_flowLow := flowLow;
prev_ackBtn  := ackBtn;

END_FUNCTION_BLOCK

(* ---- self-hard-01.raw_candidate_02.st ---- *)
FUNCTION_BLOCK FB
VAR_INPUT
    flowLow   : BOOL;
    ackBtn    : BOOL;
    sensorOK  : BOOL;
END_VAR
VAR_OUTPUT
    alarmActive : BOOL;
    alarmAcked  : BOOL;
    highHigh    : BOOL;
END_VAR
VAR
    prev_flowLow : BOOL := FALSE;
    tmp_flowRising : BOOL;
    tmp_ackRising  : BOOL;
END_VAR

(*
ENGINEERING_CONTRACT:
================================================================================
| Output/State        | Activation          | Retention      | Reset/Deact         | Scan Priority | Units/Range       |
|---------------------|---------------------|----------------|---------------------|---------------|-------------------|
| alarmActive [BOOL]  | flowLow rising edge | Until explicit | rising(ackBtn)+!flowLow+tmp_unacked_wait| Same-scan | 0..1 |
|                     |                     | deactivation   | tmp_unacked_wait:=TRUE on flowLow fall  |               |                   |
|                     |                     |                | while !alarmAcked                         |               |                   |
| alarmAcked [BOOL]   | rising(ackBtn) with | Cleared on new | rising(ackBtn)+!flowLow+tmp_unacked_wait | Same-scan | 0..1 |
|                     | flowLow present;    | flowLow rise;  |                                             |               |                   |
|                     | flowLow fall while  | retained during|                                             |               |                   |
|                     | !alarmAcked         | waiting state  |                                             |               |                   |
| highHigh [BOOL]     | !sensorOK (PUB027)  | Retained while | sensorOK TRUE (PUB035)                     | Same-scan | 0..1 |
|                     |                     | !sensorOK      |                                             |               |                   |
| tmp_unacked_wait    | flowLow falling     | Until rising   | rising(ackBtn)+!flowLow                  | Internal  | Named boolean     |
| [BOOL, local]       | while !alarmAcked   | (ackBtn)       |                                             |           |                   |
================================================================================
PUB IDs: alarmActive→PUB001/PUB002/PUB003/PUB004/PUB005/PUB006; alarmAcked→PUB007/PUB008/PUB009/PUB010/PUB011/PUB012; highHigh→PUB027/PUB035

CONTRACT_RULES: []
================================================================================
*)

tmp_flowRising := flowLow AND NOT prev_flowLow;
tmp_ackRising  := ackBtn  AND NOT prev_ackBtn;

IF tmp_flowRising THEN
    alarmActive := TRUE;
    alarmAcked  := FALSE;
ELSIF alarmActive AND tmp_ackRising THEN
    IF NOT flowLow THEN
        alarmActive := FALSE;
        alarmAcked  := FALSE;
    ELSE
        alarmAcked  := TRUE;
    END_IF;
ELSIF alarmActive AND NOT flowLow AND NOT alarmAcked AND prev_flowLow THEN
    alarmAcked := TRUE;
ELSIF alarmActive AND flowLow AND alarmAcked AND tmp_flowRising THEN
    alarmAcked := FALSE;
END_IF;

highHigh := NOT sensorOK;

prev_flowLow := flowLow;
prev_ackBtn  := ackBtn;

END_FUNCTION_BLOCK

(* ---- self-hard-01.raw_candidate_03.st ---- *)
FUNCTION_BLOCK FB
VAR_INPUT
    flowLow   : BOOL;
    ackBtn    : BOOL;
    sensorOK  : BOOL;
END_VAR
VAR_OUTPUT
    alarmActive : BOOL;
    alarmAcked  : BOOL;
    highHigh    : BOOL;
END_VAR
VAR
    prev_flowLow : BOOL := FALSE;
    prev_ackBtn  : BOOL := FALSE;
    tmp_flowRising : BOOL;
    tmp_ackRising  : BOOL;
END_VAR

(*
ENGINEERING_CONTRACT:
================================================================================
| Output/State        | Activation          | Retention      | Reset/Deact         | Scan Priority | Units/Range       |
|---------------------|---------------------|----------------|---------------------|---------------|-------------------|
| alarmActive [BOOL]  | flowLow rising edge | Until explicit | rising(ackBtn)+!flowLow; or flowLow | Same-scan | 0..1 |
|                     | (PUB001)            | deactivation   | rises while alarmAcked=TRUE (new occ) |          |                   |
| alarmAcked [BOOL]   | rising(ackBtn) with | Cleared on new | rising(ackBtn)+!flowLow (PUB009/PUB010) | Same-scan | 0..1 |
|                     | flowLow present     | flowLow rise   |                                         |               |                   |
|                     | (PUB008/PUB011);    | (new occ)      |                                         |               |                   |
|                     | flowLow falling     | Retained while |                                         |               |                   |
|                     | while !alarmAcked   | waiting clear  |                                         |               |                   |
|                     | (PUB006: pending)   | (PUB006)       |                                         |               |                   |
| highHigh [BOOL]     | !sensorOK (PUB027)  | Retained while | sensorOK TRUE (PUB035)                  | Same-scan | 0..1 |
|                     |                     | !sensorOK      |                                         |               |                   |
================================================================================
PUB IDs: alarmActive→PUB001/PUB002/PUB003/PUB004/PUB005/PUB006;
         alarmAcked→PUB006/PUB007/PUB008/PUB009/PUB010/PUB011/PUB012;
         highHigh→PUB027/PUB035

CONTRACT_RULES: []
================================================================================
*)

tmp_flowRising := flowLow AND NOT prev_flowLow;
tmp_ackRising  := ackBtn  AND NOT prev_ackBtn;

IF tmp_flowRising THEN
    alarmActive := TRUE;
    alarmAcked  := FALSE;
ELSIF alarmActive AND tmp_ackRising THEN
    IF NOT flowLow THEN
        alarmActive := FALSE;
        alarmAcked  := FALSE;
    ELSE
        alarmAcked  := TRUE;
    END_IF;
ELSIF alarmActive AND NOT flowLow AND NOT alarmAcked THEN
    alarmAcked := TRUE;
ELSIF alarmActive AND NOT flowLow AND alarmAcked THEN
    alarmActive := FALSE;
    alarmAcked  := FALSE;
END_IF;

highHigh := NOT sensorOK;

prev_flowLow := flowLow;
prev_ackBtn  := ackBtn;

END_FUNCTION_BLOCK

(* ---- self-hard-01.raw_candidate_04.st ---- *)
FUNCTION_BLOCK FB
VAR_INPUT
    flowLow   : BOOL;
    ackBtn    : BOOL;
    sensorOK  : BOOL;
END_VAR
VAR_OUTPUT
    alarmActive : BOOL;
    alarmAcked  : BOOL;
    highHigh    : BOOL;
END_VAR
VAR
    prev_flowLow : BOOL := FALSE;
    prev_ackBtn  : BOOL := FALSE;
    tmp_flowRising : BOOL;
    tmp_ackRising  : BOOL;
END_VAR

(*
ENGINEERING_CONTRACT:
================================================================================
| Output/State        | Activation          | Retention      | Reset/Deact         | Scan Priority | Units/Range       |
|---------------------|---------------------|----------------|---------------------|---------------|-------------------|
| alarmActive [BOOL]  | flowLow rising edge | Until explicit | rising(ackBtn)+!flowLow; or flowLow | Same-scan | 0..1 |
|                     | (PUB001)            | deactivation   | rises while alarmAcked=TRUE (new occ) |          |                   |
| alarmAcked [BOOL]   | rising(ackBtn) with | Cleared on new | rising(ackBtn)+!flowLow (PUB009/PUB010) | Same-scan | 0..1 |
|                     | flowLow present     | flowLow rise   |                                         |               |                   |
|                     | (PUB008/PUB011);    | (new occ)      |                                         |               |                   |
|                     | flowLow falling     | Retained while |                                         |               |                   |
|                     | while !alarmAcked   | waiting clear  |                                         |               |                   |
|                     | (PUB006: pending)   | (PUB006)       |                                         |               |                   |
| highHigh [BOOL]     | !sensorOK (PUB027)  | Retained while | sensorOK TRUE (PUB035)                  | Same-scan | 0..1 |
|                     |                     | !sensorOK      |                                         |               |                   |
================================================================================
PUB IDs: alarmActive→PUB001/PUB002/PUB003/PUB004/PUB005/PUB006;
         alarmAcked→PUB006/PUB007/PUB008/PUB009/PUB010/PUB011/PUB012;
         highHigh→PUB027/PUB035

CONTRACT_RULES: []
================================================================================
*)

tmp_flowRising := flowLow AND NOT prev_flowLow;
tmp_ackRising  := ackBtn  AND NOT prev_ackBtn;

IF tmp_flowRising THEN
    alarmActive := TRUE;
    alarmAcked  := FALSE;
ELSIF alarmActive AND tmp_ackRising AND (flowLow OR alarmAcked) THEN
    alarmAcked := TRUE;
ELSIF alarmActive AND NOT flowLow AND NOT alarmAcked THEN
    alarmAcked := TRUE;
ELSIF alarmActive AND NOT flowLow THEN
    alarmActive := FALSE;
    alarmAcked  := FALSE;
END_IF;

highHigh := NOT sensorOK;

prev_flowLow := flowLow;
prev_ackBtn  := ackBtn;

END_FUNCTION_BLOCK

(* ---- self-hard-02.candidate_01.st ---- *)
FUNCTION_BLOCK FB
VAR_INPUT
    startBtn    : BOOL;
    abortBtn    : BOOL;
    setpoint    : REAL;
    pv          : REAL;
    maxDuration : INT;
END_VAR
VAR_OUTPUT
    elapsed : INT := 0;
    phase   : INT := 0;
    timeout : BOOL := FALSE;
END_VAR
VAR
    prevStartBtn : BOOL := FALSE;
END_VAR
(* ENGINEERING_CONTRACT
+-----------------------------------------------------------+-----------------------------------+-----------------------------------+-------------------+------------+
| Output/State    | Activation              | Retention           | Explicit Reset        | Same-scan Priority | Units/Range |
+-----------------------------------------------------------+-----------------------------------+-----------------------------------+-------------------+------------+
| phase=9         | abortBtn=TRUE           | Hold until new start| New rising(startBtn)  | 1-Highest (abort)  | Enum {0,1,2,3,9} |
| phase=1         | Rising(startBtn) & no abort | Clear elapsed,timeout | Rising(startBtn)     | 2-Medium (start)   | Enum {0,1,2,3,9} |
| phase=3         | elapsed>=maxDuration    | Hold until new start| New rising(startBtn)  | 3-Lowest (running) | Enum {0,1,2,3,9} |
| elapsed         | +1 per scan when prev(1|2) | Hold in phase 3,9  | Clear on new start    | -                  | INT [0,2147483647] |
| timeout         | Set when elapsed>=maxDuration | Hold in phase 3,9 | Clear on new start   | -                  | BOOL |
+-----------------------------------------------------------+-----------------------------------+-----------------------------------+-------------------+------------+
PUB: [PUB001,PUB002,PUB003,PUB004,PUB005,PUB006,PUB007,PUB008,PUB009,PUB010,
      PUB011,PUB012,PUB013,PUB014,PUB015,PUB016,PUB017,PUB018,PUB019,PUB020,
      PUB021,PUB022,PUB023,PUB024,PUB025,PUB026,PUB027,PUB028,PUB029,PUB030,
      PUB031,PUB032,PUB033,PUB034,PUB035,PUB036,PUB037,PUB038,PUB039,PUB040,
      PUB041,PUB042,PUB043,PUB044,PUB045,PUB046,PUB047,PUB048]
*)
VAR
    tmpRisingStart : BOOL;
    tmpPrevPhase   : INT;
END_VAR

tmpRisingStart := startBtn AND NOT prevStartBtn;
tmpPrevPhase   := phase;

IF abortBtn THEN
    phase   := 9;
    elapsed := elapsed;
    timeout := timeout;
ELSIF tmpRisingStart THEN
    elapsed := 0;
    timeout := FALSE;
    phase   := 1;
ELSE
    IF (tmpPrevPhase = 1) OR (tmpPrevPhase = 2) THEN
        elapsed := elapsed + 1;
        IF elapsed >= maxDuration THEN
            timeout := TRUE;
            phase   := 3;
        ELSIF tmpPrevPhase = 1 THEN
            IF pv >= setpoint THEN
                phase := 2;
            ELSE
                phase := 1;
            END_IF;
        ELSE
            phase := 2;
        END_IF;
    ELSE
        phase := tmpPrevPhase;
    END_IF;
END_IF;

prevStartBtn := startBtn;
END_FUNCTION_BLOCK
(* CONTRACT_RULES [] *)

(* ---- self-hard-02.raw_candidate_01.st ---- *)
FUNCTION_BLOCK FB
VAR_INPUT
    startBtn    : BOOL;
    abortBtn    : BOOL;
    setpoint    : REAL;
    pv          : REAL;
    maxDuration : INT;
END_VAR
VAR_OUTPUT
    elapsed : INT := 0;
    phase   : INT := 0;
    timeout : BOOL := FALSE;
END_VAR
VAR
    prevStartBtn : BOOL := FALSE;
END_VAR
(* ENGINEERING_CONTRACT
+-----------------------------------------------------------+-----------------------------------+-----------------------------------+-------------------+------------+
| Output/State    | Activation              | Retention           | Explicit Reset        | Same-scan Priority | Units/Range |
+-----------------------------------------------------------+-----------------------------------+-----------------------------------+-------------------+------------+
| phase=9         | abortBtn=TRUE           | Hold until new start| New rising(startBtn)  | 1-Highest (abort)  | Enum {0,1,2,3,9} |
| phase=1         | Rising(startBtn) & no abort | Clear elapsed,timeout | Rising(startBtn)     | 2-Medium (start)   | Enum {0,1,2,3,9} |
| phase=3         | elapsed>=maxDuration    | Hold until new start| New rising(startBtn)  | 3-Lowest (running) | Enum {0,1,2,3,9} |
| elapsed         | +1 per scan when prev(1|2) | Hold in phase 3,9  | Clear on new start    | -                  | INT [0,2147483647] |
| timeout         | Set when elapsed>=maxDuration | Hold in phase 3,9 | Clear on new start   | -                  | BOOL |
+-----------------------------------------------------------+-----------------------------------+-----------------------------------+-------------------+------------+
PUB: [PUB001,PUB002,PUB003,PUB004,PUB005,PUB006,PUB007,PUB008,PUB009,PUB010,
      PUB011,PUB012,PUB013,PUB014,PUB015,PUB016,PUB017,PUB018,PUB019,PUB020,
      PUB021,PUB022,PUB023,PUB024,PUB025,PUB026,PUB027,PUB028,PUB029,PUB030,
      PUB031,PUB032,PUB033,PUB034,PUB035,PUB036,PUB037,PUB038,PUB039,PUB040,
      PUB041,PUB042,PUB043,PUB044,PUB045,PUB046,PUB047,PUB048]
*)
VAR
    tmpRisingStart : BOOL;
    tmpPrevPhase   : INT;
END_VAR

tmpRisingStart := startBtn AND NOT prevStartBtn;
tmpPrevPhase   := phase;

IF abortBtn THEN
    phase   := 9;
    elapsed := elapsed;
    timeout := timeout;
ELSIF tmpRisingStart THEN
    elapsed := 0;
    timeout := FALSE;
    phase   := 1;
ELSE
    IF (tmpPrevPhase = 1) OR (tmpPrevPhase = 2) THEN
        elapsed := elapsed + 1;
        IF elapsed >= maxDuration THEN
            timeout := TRUE;
            phase   := 3;
        ELSIF tmpPrevPhase = 1 THEN
            IF pv >= setpoint THEN
                phase := 2;
            ELSE
                phase := 1;
            END_IF;
        ELSE
            phase := 2;
        END_IF;
    ELSE
        phase := tmpPrevPhase;
    END_IF;
END_IF;

prevStartBtn := startBtn;
END_FUNCTION_BLOCK
(* CONTRACT_RULES [] *)

(* ---- self-hard-03.candidate_02.st ---- *)
(* ENGINEERING_CONTRACT
| Output/State    | Activation        | Retention         | Explicit Reset | Scan Priority | Units/Boundaries |
|-----------------|-------------------|-------------------|----------------|---------------|------------------|
| count           | Computed each scan| Maintained        | None           | After ops     | 0..8 integer     |
| full            | count=8           | Held until count<8| None           | With count    | BOOL             |
| empty           | count=0           | Held until count>0| None           | With count    | BOOL             |
| head            | fifo[1] or 0      | Held on empty     | None           | After ops     | INT              |
| fifo[1..count]  | Compacted each scan| Retained         | None           | After ops     | ARRAY[1..8] INT  |

PUB001: pushEn (rising edge trigger)
PUB002: pushItem (INT payload)
PUB003: popEn (rising edge trigger)
PUB004: fifo INOUT ARRAY[1..8] INT, caller-bound, read-write during scan
PUB005: count = length 0..8
PUB006: full <-> count=8
PUB007: empty <-> count=0
PUB008: head = fifo[1] when !empty else 0
PUB009: pop on rising(popEn) executes first if count>0
PUB010: push on rising(pushEn) executes second if count<8
PUB011: same-scan full+pop+push: pop frees slot then push appends
PUB012: same-scan empty+pop+push: only push adds item
PUB013: fifo[1..count] compact, fifo[1]=head when !empty
PUB014: undefined fifo[count+1..8]
PUB015: initial count=0, empty=TRUE, fifo[1..8] undefined
PUB016: rising edge = prev=FALSE AND cur=TRUE
PUB017: sustained press does not repeat (edge-only)
PUB018: R_TRIG used for edge memory
PUB019: scan-order: detect edges, execute pop, execute push, compute outputs
PUB020: CONTRACT_RULES []
*)
FUNCTION_BLOCK FB
VAR_INPUT
    pushEn : BOOL;
    pushItem : INT;
    popEn : BOOL;
END_VAR
VAR_IN_OUT
    fifo : ARRAY[1..8] OF INT;
END_VAR
VAR_OUTPUT
    count : INT := 0;
    full : BOOL := FALSE;
    empty : BOOL := TRUE;
    head : INT := 0;
END_VAR
VAR
    pushTrig : R_TRIG;
    popTrig : R_TRIG;
    i : INT;
END_VAR

pushTrig(CLK := pushEn);
popTrig(CLK := popEn);

IF popTrig.Q AND count > 0 THEN
    FOR i := 1 TO count - 1 DO
        fifo[i] := fifo[i + 1];
    END_FOR;
    count := count - 1;
END_IF;

IF pushTrig.Q AND count < 8 THEN
    count := count + 1;
    fifo[count] := pushItem;
END_IF;

full := (count = 8);
empty := (count = 0);
head := 0;
IF NOT empty THEN
    head := fifo[1];
END_IF;

END_FUNCTION_BLOCK

(* ---- self-hard-03.raw_candidate_02.st ---- *)
(* ENGINEERING_CONTRACT
| Output/State    | Activation        | Retention         | Explicit Reset | Scan Priority | Units/Boundaries |
|-----------------|-------------------|-------------------|----------------|---------------|------------------|
| count           | Computed each scan| Maintained        | None           | After ops     | 0..8 integer     |
| full            | count=8           | Held until count<8| None           | With count    | BOOL             |
| empty           | count=0           | Held until count>0| None           | With count    | BOOL             |
| head            | fifo[1] or 0      | Held on empty     | None           | After ops     | INT              |
| fifo[1..count]  | Compacted each scan| Retained         | None           | After ops     | ARRAY[1..8] INT  |

PUB001: pushEn (rising edge trigger)
PUB002: pushItem (INT payload)
PUB003: popEn (rising edge trigger)
PUB004: fifo INOUT ARRAY[1..8] INT, caller-bound, read-write during scan
PUB005: count = length 0..8
PUB006: full <-> count=8
PUB007: empty <-> count=0
PUB008: head = fifo[1] when !empty else 0
PUB009: pop on rising(popEn) executes first if count>0
PUB010: push on rising(pushEn) executes second if count<8
PUB011: same-scan full+pop+push: pop frees slot then push appends
PUB012: same-scan empty+pop+push: only push adds item
PUB013: fifo[1..count] compact, fifo[1]=head when !empty
PUB014: undefined fifo[count+1..8]
PUB015: initial count=0, empty=TRUE, fifo[1..8] undefined
PUB016: rising edge = prev=FALSE AND cur=TRUE
PUB017: sustained press does not repeat (edge-only)
PUB018: R_TRIG used for edge memory
PUB019: scan-order: detect edges, execute pop, execute push, compute outputs
PUB020: CONTRACT_RULES []
*)
FUNCTION_BLOCK FB
VAR_INPUT
    pushEn : BOOL;
    pushItem : INT;
    popEn : BOOL;
END_VAR
VAR_IN_OUT
    fifo : ARRAY[1..8] OF INT;
END_VAR
VAR_OUTPUT
    count : INT := 0;
    full : BOOL := FALSE;
    empty : BOOL := TRUE;
    head : INT := 0;
END_VAR
VAR
    pushTrig : R_TRIG;
    popTrig : R_TRIG;
    i : INT;
END_VAR

pushTrig(CLK := pushEn);
popTrig(CLK := popEn);

IF popTrig.Q AND count > 0 THEN
    FOR i := 1 TO count - 1 DO
        fifo[i] := fifo[i + 1];
    END_FOR;
    count := count - 1;
END_IF;

IF pushTrig.Q AND count < 8 THEN
    count := count + 1;
    fifo[count] := pushItem;
END_IF;

full := (count = 8);
empty := (count = 0);
head := 0;
IF NOT empty THEN
    head := fifo[1];
END_IF;

END_FUNCTION_BLOCK

(* ---- self-hard-04.candidate_01.st ---- *)
FUNCTION_BLOCK FB
VAR_OUTPUT
    leadPump : INT := 0;
    lagPump : INT := 0;
    runningCount : INT := 0;
END_VAR
VAR_INPUT
    demand : INT;
    runHours : ARRAY[1..5] OF LINT;
    rotated : BOOL;
END_VAR
VAR
    prevLeadPump : INT := 0;
    prevLagPump : INT := 0;
    prevRunningCount : INT := 0;
    tmpLead : INT;
    tmpLag : INT;
    tmpCount : INT;
    minHours : LINT;
    minPump : INT;
    i : INT;
END_VAR
VAR_TEMP
    local_i : INT;
END_VAR
(*
ENGINEERING_CONTRACT:
| State Group         | Activation           | Retention/Hold           | Explicit Reset         | Same-Scan Priority | Units/Boundaries         |
|---------------------|----------------------|--------------------------|------------------------|--------------------|--------------------------|
| runningCount [S1]   | demand>0             | hold value               | demand<=0→0            | same-scan assign   | 0..5 (clipped from demand)|
| leadPump [S2,S3]    | demand>0, prevLead=0 | hold during positive dem | demand<=0→0            | initial selection first | 0 or 1..5                |
| leadPump rotation   | rotated=TRUE AND >50h diff | hold until next valid trigger | demand<=0→0 | rotation evaluated after initial | 1..5 only               |
| lagPump [S2,S8,S9]  | demand>=2 AND (initial/change/rise) | hold when unchanged | demand<=1→0           | evaluated after lead | 0 or 1..5, ≠leadPump     |
PUB clauses: PUB001(s0), PUB002(demand), PUB003(clipped), PUB004(ascending), PUB005(different), PUB006(0→pos), PUB007(hysteresis50h), PUB008(level-rotated), PUB009(no req→no change), PUB010(demand=0→clr), PUB011(lag selection moments), PUB012(no reselection), PUB013(index 1..5)
*)
(* CONTRACT_RULES [] *)

tmpLead := prevLeadPump;
tmpLag := prevLagPump;
tmpCount := prevRunningCount;

tmpCount := demand;
IF demand < 0 THEN
    tmpCount := 0;
END_IF;
IF demand > 5 THEN
    tmpCount := 5;
END_IF;

IF demand <= 0 THEN
    tmpLead := 0;
    tmpLag := 0;
ELSIF tmpLead = 0 THEN
    minHours := runHours[1];
    minPump := 1;
    FOR local_i := 2 TO 5 DO
        IF runHours[local_i] < minHours OR (runHours[local_i] = minHours AND local_i < minPump) THEN
            minHours := runHours[local_i];
            minPump := local_i;
        END_IF;
    END_FOR;
    tmpLead := minPump;
    IF tmpCount >= 2 THEN
        minHours := LINT#16#7FFFFFFFFFFFFFFF;
        minPump := 0;
        FOR local_i := 1 TO 5 DO
            IF local_i <> tmpLead THEN
                IF runHours[local_i] < minHours OR (runHours[local_i] = minHours AND local_i < minPump) THEN
                    minHours := runHours[local_i];
                    minPump := local_i;
                END_IF;
            END_IF;
        END_FOR;
        tmpLag := minPump;
    ELSE
        tmpLag := 0;
    END_IF;
ELSE
    IF rotated THEN
        minHours := runHours[1];
        minPump := 1;
        FOR local_i := 2 TO 5 DO
            IF runHours[local_i] < minHours OR (runHours[local_i] = minHours AND local_i < minPump) THEN
                minHours := runHours[local_i];
                minPump := local_i;
            END_IF;
        END_FOR;
        IF runHours[tmpLead] > minHours + LINT#50 THEN
            tmpLead := minPump;
        END_IF;
    END_IF;
    IF tmpCount >= 2 THEN
        IF tmpLead <> prevLeadPump OR tmpCount > prevRunningCount THEN
            minHours := LINT#16#7FFFFFFFFFFFFFFF;
            minPump := 0;
            FOR local_i := 1 TO 5 DO
                IF local_i <> tmpLead THEN
                    IF runHours[local_i] < minHours OR (runHours[local_i] = minHours AND local_i < minPump) THEN
                        minHours := runHours[local_i];
                        minPump := local_i;
                    END_IF;
                END_IF;
            END_FOR;
            tmpLag := minPump;
        END_IF;
    ELSE
        tmpLag := 0;
    END_IF;
END_IF;

leadPump := tmpLead;
lagPump := tmpLag;
runningCount := tmpCount;
prevLeadPump := tmpLead;
prevLagPump := tmpLag;
prevRunningCount := tmpCount;
END_FUNCTION_BLOCK

(* ---- self-hard-04.raw_candidate_01.st ---- *)
FUNCTION_BLOCK FB
VAR_OUTPUT
    leadPump : INT := 0;
    lagPump : INT := 0;
    runningCount : INT := 0;
END_VAR
VAR_INPUT
    demand : INT;
    runHours : ARRAY[1..5] OF LINT;
    rotated : BOOL;
END_VAR
VAR
    prevLeadPump : INT := 0;
    prevLagPump : INT := 0;
    prevRunningCount : INT := 0;
    tmpLead : INT;
    tmpLag : INT;
    tmpCount : INT;
    minHours : LINT;
    minPump : INT;
    i : INT;
END_VAR
VAR_TEMP
    local_i : INT;
END_VAR
(*
ENGINEERING_CONTRACT:
| State Group         | Activation           | Retention/Hold           | Explicit Reset         | Same-Scan Priority | Units/Boundaries         |
|---------------------|----------------------|--------------------------|------------------------|--------------------|--------------------------|
| runningCount [S1]   | demand>0             | hold value               | demand<=0→0            | same-scan assign   | 0..5 (clipped from demand)|
| leadPump [S2,S3]    | demand>0, prevLead=0 | hold during positive dem | demand<=0→0            | initial selection first | 0 or 1..5                |
| leadPump rotation   | rotated=TRUE AND >50h diff | hold until next valid trigger | demand<=0→0 | rotation evaluated after initial | 1..5 only               |
| lagPump [S2,S8,S9]  | demand>=2 AND (initial/change/rise) | hold when unchanged | demand<=1→0           | evaluated after lead | 0 or 1..5, ≠leadPump     |
PUB clauses: PUB001(s0), PUB002(demand), PUB003(clipped), PUB004(ascending), PUB005(different), PUB006(0→pos), PUB007(hysteresis50h), PUB008(level-rotated), PUB009(no req→no change), PUB010(demand=0→clr), PUB011(lag selection moments), PUB012(no reselection), PUB013(index 1..5)
*)
(* CONTRACT_RULES [] *)

tmpLead := prevLeadPump;
tmpLag := prevLagPump;
tmpCount := prevRunningCount;

tmpCount := demand;
IF demand < 0 THEN
    tmpCount := 0;
END_IF
IF demand > 5 THEN
    tmpCount := 5;
END_IF

IF demand <= 0 THEN
    tmpLead := 0;
    tmpLag := 0;
ELSIF tmpLead = 0 THEN
    minHours := runHours[1];
    minPump := 1;
    FOR local_i := 2 TO 5 DO
        IF runHours[local_i] < minHours OR (runHours[local_i] = minHours AND local_i < minPump) THEN
            minHours := runHours[local_i];
            minPump := local_i;
        END_IF
    END_FOR
    tmpLead := minPump;
    IF tmpCount >= 2 THEN
        minHours := LINT#16#7FFFFFFFFFFFFFFF;
        minPump := 0;
        FOR local_i := 1 TO 5 DO
            IF local_i <> tmpLead THEN
                IF runHours[local_i] < minHours OR (runHours[local_i] = minHours AND local_i < minPump) THEN
                    minHours := runHours[local_i];
                    minPump := local_i;
                END_IF
            END_IF
        END_FOR
        tmpLag := minPump;
    ELSE
        tmpLag := 0;
    END_IF
ELSE
    IF rotated THEN
        minHours := runHours[1];
        minPump := 1;
        FOR local_i := 2 TO 5 DO
            IF runHours[local_i] < minHours OR (runHours[local_i] = minHours AND local_i < minPump) THEN
                minHours := runHours[local_i];
                minPump := local_i;
            END_IF
        END_FOR
        IF runHours[tmpLead] > minHours + LINT#50 THEN
            tmpLead := minPump;
        END_IF
    END_IF
    IF tmpCount >= 2 THEN
        IF tmpLead <> prevLeadPump OR tmpCount > prevRunningCount THEN
            minHours := LINT#16#7FFFFFFFFFFFFFFF;
            minPump := 0;
            FOR local_i := 1 TO 5 DO
                IF local_i <> tmpLead THEN
                    IF runHours[local_i] < minHours OR (runHours[local_i] = minHours AND local_i < minPump) THEN
                        minHours := runHours[local_i];
                        minPump := local_i;
                    END_IF
                END_IF
            END_FOR
            tmpLag := minPump;
        END_IF
    ELSE
        tmpLag := 0;
    END_IF
END_IF

leadPump := tmpLead;
lagPump := tmpLag;
runningCount := tmpCount;
prevLeadPump := tmpLead;
prevLagPump := tmpLag;
prevRunningCount := tmpCount;
END_FUNCTION_BLOCK

(* ---- self-hard-05.candidate_01.st ---- *)
FUNCTION_BLOCK FB
VAR_INPUT
    runRequest  : BOOL;
    flameOK     : BOOL;
    o2Valid     : BOOL;
    o2PV        : REAL;
    baseAir     : REAL;
    resetBtn    : BOOL;
END_VAR
VAR_OUTPUT
    fuelPermit  : BOOL;
    trimEnable  : BOOL;
    airTrim     : REAL;
    airCommand  : REAL;
    tripLatched : BOOL;
    o2Fault     : BOOL;
END_VAR
VAR
    prev_resetBtn : BOOL := FALSE;
END_VAR

// ENGINEERING_CONTRACT
// [S1]  PUB003   tripLatched: ACTIVE when runRequest & !flameOK (same scan, no delay)
// [S2]  PUB008   tripLatched: HOLD until rising(resetBtn) & !runRequest & !flameOK
// [S3]  PUB008   tripLatched: inhibit fuelPermit while held (same scan)
// [S4]  PUB004   fuelPermit: ACTIVE when runRequest & flameOK & !tripLatched
// [S5]  PUB010   airCommand: FORCE 0.0 when !fuelPermit (same scan)
// [S6]  PUB010   airCommand: CLAMP [0.0, 100.0] always
// [S7]  PUB005   airTrim: CLAMP [-10.0, 10.0] always
// [S8]  PUB008   trimEnable: ACTIVE when fuelPermit & !o2Fault
// [S9]  PUB007   o2Fault: ACTIVE when !o2Valid | o2PV<0 | o2PV>21
// [S10] PUB008   airTrim: FORCE 0.0 when !trimEnable (no residual)
// [S11-S12] PUB006 airTrim: =2*(2-o2PV) raw, -10 limit only when o2PV>7
// [S13-S14] PUB010 airCommand: CLAMP [0,100] after baseAir+airTrim sum
// Reset: PUB023 edge-triggered, not level. Same-scan priority per S1/S3.

LOCAL_EDGE_TRIGGER(resetBtn, prev_resetBtn);
o2Fault := NOT o2Valid OR o2PV < 0.0 OR o2PV > 21.0;
tripLatched := tripLatched OR (runRequest AND NOT flameOK);
IF LOCAL_EDGE_TRIG_RISE AND NOT runRequest AND NOT flameOK THEN
    tripLatched := FALSE;
END_IF;
fuelPermit := runRequest AND flameOK AND NOT tripLatched;
trimEnable := fuelPermit AND NOT o2Fault;
IF trimEnable THEN
    airTrim := LIMIT(-10.0, 2.0 * (2.0 - o2PV), 10.0);
ELSE
    airTrim := 0.0;
END_IF;
IF fuelPermit THEN
    airCommand := LIMIT(0.0, baseAir + airTrim, 100.0);
ELSE
    airCommand := 0.0;
END_IF;
prev_resetBtn := resetBtn;
END_FUNCTION_BLOCK

(* CONTRACT_RULES [] *)

(* ---- self-hard-05.candidate_02.st ---- *)
FUNCTION_BLOCK FB
VAR_INPUT
    runRequest  : BOOL;
    flameOK     : BOOL;
    o2Valid     : BOOL;
    o2PV        : REAL;
    baseAir     : REAL;
    resetBtn    : BOOL;
END_VAR
VAR_OUTPUT
    fuelPermit  : BOOL;
    trimEnable  : BOOL;
    airTrim     : REAL;
    airCommand  : REAL;
    tripLatched : BOOL;
    o2Fault     : BOOL;
END_VAR
VAR
    prev_resetBtn : BOOL := FALSE;
END_VAR

// ENGINEERING_CONTRACT
// [S1]  PUB003   tripLatched: ACTIVE when runRequest & !flameOK (same scan, no delay)
// [S2]  PUB008   tripLatched: HOLD until rising(resetBtn) & !runRequest & !flameOK
// [S3]  PUB008   tripLatched: inhibit fuelPermit while held (same scan)
// [S4]  PUB004   fuelPermit: ACTIVE when runRequest & flameOK & !tripLatched
// [S5]  PUB010   airCommand: FORCE 0.0 when !fuelPermit (same scan)
// [S6]  PUB010   airCommand: CLAMP [0.0, 100.0] always
// [S7]  PUB005   airTrim: CLAMP [-10.0, 10.0] always
// [S8]  PUB008   trimEnable: ACTIVE when fuelPermit & !o2Fault
// [S9]  PUB007   o2Fault: ACTIVE when !o2Valid | o2PV<0 | o2PV>21
// [S10] PUB008   airTrim: FORCE 0.0 when !trimEnable (no residual)
// [S11-S12] PUB006 airTrim: =2*(2-o2PV) raw, -10 limit only when o2PV>7
// [S13-S14] PUB010 airCommand: CLAMP [0,100] after baseAir+airTrim sum
// Reset: PUB023 edge-triggered, not level. Same-scan priority per S1/S3.

LOCAL_EDGE_TRIG_RISE := resetBtn AND NOT prev_resetBtn;
o2Fault := NOT o2Valid OR o2PV < 0.0 OR o2PV > 21.0;
tripLatched := tripLatched OR (runRequest AND NOT flameOK);
IF LOCAL_EDGE_TRIG_RISE AND NOT runRequest AND NOT flameOK THEN
    tripLatched := FALSE;
END_IF;
fuelPermit := runRequest AND flameOK AND NOT tripLatched;
trimEnable := fuelPermit AND NOT o2Fault;
IF trimEnable THEN
    airTrim := LIMIT(-10.0, 2.0 * (2.0 - o2PV), 10.0);
ELSE
    airTrim := 0.0;
END_IF;
IF fuelPermit THEN
    airCommand := LIMIT(0.0, baseAir + airTrim, 100.0);
ELSE
    airCommand := 0.0;
END_IF;
prev_resetBtn := resetBtn;
END_FUNCTION_BLOCK

(* CONTRACT_RULES [] *)

(* ---- self-hard-05.candidate_03.st ---- *)
FUNCTION_BLOCK FB
VAR_INPUT
    runRequest  : BOOL;
    flameOK     : BOOL;
    o2Valid     : BOOL;
    o2PV        : REAL;
    baseAir     : REAL;
    resetBtn    : BOOL;
END_VAR
VAR_OUTPUT
    fuelPermit  : BOOL;
    trimEnable  : BOOL;
    airTrim     : REAL;
    airCommand  : REAL;
    tripLatched : BOOL;
    o2Fault     : BOOL;
END_VAR
VAR
    prev_resetBtn : BOOL := FALSE;
    tmp_resetRising : BOOL;
END_VAR

// ENGINEERING_CONTRACT
// [S1]  PUB003   tripLatched: ACTIVE when runRequest & !flameOK (same scan, no delay)
// [S2]  PUB008   tripLatched: HOLD until rising(resetBtn) & !runRequest & !flameOK
// [S3]  PUB008   tripLatched: inhibit fuelPermit while held (same scan)
// [S4]  PUB004   fuelPermit: ACTIVE when runRequest & flameOK & !tripLatched
// [S5]  PUB010   airCommand: FORCE 0.0 when !fuelPermit (same scan)
// [S6]  PUB010   airCommand: CLAMP [0.0, 100.0] always
// [S7]  PUB005   airTrim: CLAMP [-10.0, 10.0] always
// [S8]  PUB008   trimEnable: ACTIVE when fuelPermit & !o2Fault
// [S9]  PUB007   o2Fault: ACTIVE when !o2Valid | o2PV<0 | o2PV>21
// [S10] PUB008   airTrim: FORCE 0.0 when !trimEnable (no residual)
// [S11-S12] PUB006 airTrim: =2*(2-o2PV) raw, -10 limit only when o2PV>7
// [S13-S14] PUB010 airCommand: CLAMP [0,100] after baseAir+airTrim sum
// Reset: PUB023 edge-triggered, not level. Same-scan priority per S1/S3.

tmp_resetRising := resetBtn AND NOT prev_resetBtn;
o2Fault := NOT o2Valid OR o2PV < 0.0 OR o2PV > 21.0;
tripLatched := tripLatched OR (runRequest AND NOT flameOK);
IF tmp_resetRising AND NOT runRequest AND NOT flameOK THEN
    tripLatched := FALSE;
END_IF;
fuelPermit := runRequest AND flameOK AND NOT tripLatched;
trimEnable := fuelPermit AND NOT o2Fault;
IF trimEnable THEN
    airTrim := LIMIT(-10.0, 2.0 * (2.0 - o2PV), 10.0);
ELSE
    airTrim := 0.0;
END_IF;
IF fuelPermit THEN
    airCommand := LIMIT(0.0, baseAir + airTrim, 100.0);
ELSE
    airCommand := 0.0;
END_IF;
prev_resetBtn := resetBtn;
END_FUNCTION_BLOCK

(* CONTRACT_RULES [] *)

(* ---- self-hard-05.raw_candidate_01.st ---- *)
FUNCTION_BLOCK FB
VAR_INPUT
    runRequest  : BOOL;
    flameOK     : BOOL;
    o2Valid     : BOOL;
    o2PV        : REAL;
    baseAir     : REAL;
    resetBtn    : BOOL;
END_VAR
VAR_OUTPUT
    fuelPermit  : BOOL;
    trimEnable  : BOOL;
    airTrim     : REAL;
    airCommand  : REAL;
    tripLatched : BOOL;
    o2Fault     : BOOL;
END_VAR
VAR
    prev_resetBtn : BOOL := FALSE;
END_VAR

// ENGINEERING_CONTRACT
// [S1]  PUB003   tripLatched: ACTIVE when runRequest & !flameOK (same scan, no delay)
// [S2]  PUB008   tripLatched: HOLD until rising(resetBtn) & !runRequest & !flameOK
// [S3]  PUB008   tripLatched: inhibit fuelPermit while held (same scan)
// [S4]  PUB004   fuelPermit: ACTIVE when runRequest & flameOK & !tripLatched
// [S5]  PUB010   airCommand: FORCE 0.0 when !fuelPermit (same scan)
// [S6]  PUB010   airCommand: CLAMP [0.0, 100.0] always
// [S7]  PUB005   airTrim: CLAMP [-10.0, 10.0] always
// [S8]  PUB008   trimEnable: ACTIVE when fuelPermit & !o2Fault
// [S9]  PUB007   o2Fault: ACTIVE when !o2Valid | o2PV<0 | o2PV>21
// [S10] PUB008   airTrim: FORCE 0.0 when !trimEnable (no residual)
// [S11-S12] PUB006 airTrim: =2*(2-o2PV) raw, -10 limit only when o2PV>7
// [S13-S14] PUB010 airCommand: CLAMP [0,100] after baseAir+airTrim sum
// Reset: PUB023 edge-triggered, not level. Same-scan priority per S1/S3.

LOCAL_EDGE_TRIGGER(resetBtn, prev_resetBtn);
o2Fault := NOT o2Valid OR o2PV < 0.0 OR o2PV > 21.0;
tripLatched := tripLatched OR (runRequest AND NOT flameOK);
IF LOCAL_EDGE_TRIG_RISE AND NOT runRequest AND NOT flameOK THEN
    tripLatched := FALSE;
END_IF;
fuelPermit := runRequest AND flameOK AND NOT tripLatched;
trimEnable := fuelPermit AND NOT o2Fault;
IF trimEnable THEN
    airTrim := LIMIT(-10.0, 2.0 * (2.0 - o2PV), 10.0);
ELSE
    airTrim := 0.0;
END_IF;
IF fuelPermit THEN
    airCommand := LIMIT(0.0, baseAir + airTrim, 100.0);
ELSE
    airCommand := 0.0;
END_IF;
prev_resetBtn := resetBtn;
END_FUNCTION_BLOCK

(* CONTRACT_RULES [] *)

(* ---- self-hard-05.raw_candidate_02.st ---- *)
FUNCTION_BLOCK FB
VAR_INPUT
    runRequest  : BOOL;
    flameOK     : BOOL;
    o2Valid     : BOOL;
    o2PV        : REAL;
    baseAir     : REAL;
    resetBtn    : BOOL;
END_VAR
VAR_OUTPUT
    fuelPermit  : BOOL;
    trimEnable  : BOOL;
    airTrim     : REAL;
    airCommand  : REAL;
    tripLatched : BOOL;
    o2Fault     : BOOL;
END_VAR
VAR
    prev_resetBtn : BOOL := FALSE;
END_VAR

// ENGINEERING_CONTRACT
// [S1]  PUB003   tripLatched: ACTIVE when runRequest & !flameOK (same scan, no delay)
// [S2]  PUB008   tripLatched: HOLD until rising(resetBtn) & !runRequest & !flameOK
// [S3]  PUB008   tripLatched: inhibit fuelPermit while held (same scan)
// [S4]  PUB004   fuelPermit: ACTIVE when runRequest & flameOK & !tripLatched
// [S5]  PUB010   airCommand: FORCE 0.0 when !fuelPermit (same scan)
// [S6]  PUB010   airCommand: CLAMP [0.0, 100.0] always
// [S7]  PUB005   airTrim: CLAMP [-10.0, 10.0] always
// [S8]  PUB008   trimEnable: ACTIVE when fuelPermit & !o2Fault
// [S9]  PUB007   o2Fault: ACTIVE when !o2Valid | o2PV<0 | o2PV>21
// [S10] PUB008   airTrim: FORCE 0.0 when !trimEnable (no residual)
// [S11-S12] PUB006 airTrim: =2*(2-o2PV) raw, -10 limit only when o2PV>7
// [S13-S14] PUB010 airCommand: CLAMP [0,100] after baseAir+airTrim sum
// Reset: PUB023 edge-triggered, not level. Same-scan priority per S1/S3.

LOCAL_EDGE_TRIG_RISE := resetBtn AND NOT prev_resetBtn;
o2Fault := NOT o2Valid OR o2PV < 0.0 OR o2PV > 21.0;
tripLatched := tripLatched OR (runRequest AND NOT flameOK);
IF LOCAL_EDGE_TRIG_RISE AND NOT runRequest AND NOT flameOK THEN
    tripLatched := FALSE;
END_IF;
fuelPermit := runRequest AND flameOK AND NOT tripLatched;
trimEnable := fuelPermit AND NOT o2Fault;
IF trimEnable THEN
    airTrim := LIMIT(-10.0, 2.0 * (2.0 - o2PV), 10.0);
ELSE
    airTrim := 0.0;
END_IF;
IF fuelPermit THEN
    airCommand := LIMIT(0.0, baseAir + airTrim, 100.0);
ELSE
    airCommand := 0.0;
END_IF;
prev_resetBtn := resetBtn;
END_FUNCTION_BLOCK

(* CONTRACT_RULES [] *)

(* ---- self-hard-05.raw_candidate_03.st ---- *)
FUNCTION_BLOCK FB
VAR_INPUT
    runRequest  : BOOL;
    flameOK     : BOOL;
    o2Valid     : BOOL;
    o2PV        : REAL;
    baseAir     : REAL;
    resetBtn    : BOOL;
END_VAR
VAR_OUTPUT
    fuelPermit  : BOOL;
    trimEnable  : BOOL;
    airTrim     : REAL;
    airCommand  : REAL;
    tripLatched : BOOL;
    o2Fault     : BOOL;
END_VAR
VAR
    prev_resetBtn : BOOL := FALSE;
    tmp_resetRising : BOOL;
END_VAR

// ENGINEERING_CONTRACT
// [S1]  PUB003   tripLatched: ACTIVE when runRequest & !flameOK (same scan, no delay)
// [S2]  PUB008   tripLatched: HOLD until rising(resetBtn) & !runRequest & !flameOK
// [S3]  PUB008   tripLatched: inhibit fuelPermit while held (same scan)
// [S4]  PUB004   fuelPermit: ACTIVE when runRequest & flameOK & !tripLatched
// [S5]  PUB010   airCommand: FORCE 0.0 when !fuelPermit (same scan)
// [S6]  PUB010   airCommand: CLAMP [0.0, 100.0] always
// [S7]  PUB005   airTrim: CLAMP [-10.0, 10.0] always
// [S8]  PUB008   trimEnable: ACTIVE when fuelPermit & !o2Fault
// [S9]  PUB007   o2Fault: ACTIVE when !o2Valid | o2PV<0 | o2PV>21
// [S10] PUB008   airTrim: FORCE 0.0 when !trimEnable (no residual)
// [S11-S12] PUB006 airTrim: =2*(2-o2PV) raw, -10 limit only when o2PV>7
// [S13-S14] PUB010 airCommand: CLAMP [0,100] after baseAir+airTrim sum
// Reset: PUB023 edge-triggered, not level. Same-scan priority per S1/S3.

tmp_resetRising := resetBtn AND NOT prev_resetBtn;
o2Fault := NOT o2Valid OR o2PV < 0.0 OR o2PV > 21.0;
tripLatched := tripLatched OR (runRequest AND NOT flameOK);
IF tmp_resetRising AND NOT runRequest AND NOT flameOK THEN
    tripLatched := FALSE;
END_IF;
fuelPermit := runRequest AND flameOK AND NOT tripLatched;
trimEnable := fuelPermit AND NOT o2Fault;
IF trimEnable THEN
    airTrim := LIMIT(-10.0, 2.0 * (2.0 - o2PV), 10.0);
ELSE
    airTrim := 0.0;
END_IF;
IF fuelPermit THEN
    airCommand := LIMIT(0.0, baseAir + airTrim, 100.0);
ELSE
    airCommand := 0.0;
END_IF;
prev_resetBtn := resetBtn;
END_FUNCTION_BLOCK

(* CONTRACT_RULES [] *)

(* ---- self-hard-06.candidate_01.st ---- *)
FUNCTION_BLOCK FB
VAR_INPUT
    runRequest      : BOOL;
    pressure        : REAL;
    pressureValid   : BOOL;
    fuelFlow        : REAL;
    steamFlow       : REAL;
    outletCmd       : INT;
    outletFeedback  : INT;
    resetBtn        : BOOL;
END_VAR
VAR_OUTPUT
    tripLatched     : BOOL;
    fuelPermit      : BOOL;
    currentCauseMask: WORD;
    latchedCauseMask: WORD;
    diagnosticActive: BOOL;
END_VAR
VAR
    prevResetBtn    : BOOL := FALSE;
    prevRunRequest  : BOOL := FALSE;
    prevPressureValid : BOOL := FALSE;
    prevPressure    : REAL := 0.0;
    prevFuelFlow    : REAL := 0.0;
    prevSteamFlow   : REAL := 0.0;
    prevOutletCmd   : INT := 0;
    prevOutletFeedback : INT := 0;
    prevTripLatched : BOOL := FALSE;
    prevCurrentCauseMask : WORD := 0;
    prevLatchedCauseMask : WORD := 0;
    stuckValveConsecutiveCount : INT := 0;
    tmpRisingReset  : BOOL;
    tmpRisingPrevCond : BOOL;
    tmpTwoAgoPrevCond : BOOL;
    tmpStuckCond   : BOOL;
    tmpCurrentMask : WORD;
    tmpOverpressureValid : BOOL;
END_VAR

(* CONTRACT:
   | Output/State    | Activation         | Retention       | Reset/Deactivation           | Same-scan Priority | Units/Boundaries       |
   |-----------------|--------------------|-----------------|-------------------------------|--------------------|------------------------|
   | tripLatched     | runRequest & (!pressureValid OR pressure>=4500.0) | Hold until resetBtn rising & !runRequest & pressureValid & pressure<=4200.0 | resetBtn rising edge clears | Same-scan with clue calc | BOOL; 4500/4200 kPa hysteresis |
   | fuelPermit      | runRequest & !tripLatched | None (combinational) | Clears when tripLatched sets | Same-scan | BOOL |
   | currentCauseMask| Recalc every scan | None (recalculated) | Zero when !runRequest | Same-scan | WORD bits 0-3; 0,1,2,4,6,8 only |
   | latchedCauseMask| OR into when tripLatched | Accumulate across trip | Clear on valid reset | Same-scan | WORD bits 0-3; 0-15 |
   | diagnosticActive| currentCauseMask <> 0 | None | Clears when mask zero | Same-scan | BOOL |
   | stuckValveConsecutiveCount | Increment when stuckCond true 3+ scans | Hold | Reset on any break in condition | Per-scan counter | INT; 0-3+ |

   PUB: PUB001(trip on !pressureValid), PUB002(overpressure>=4500), PUB003(clear hysteresis), PUB004(!runRequest=>mask=0),
        PUB005(stuck valve 3-scan), PUB006(latched accumulation), PUB007(fuelPermit), PUB008(diagnosticActive),
        PUB009(bit3 unlocated), PUB010(bit0 transmitter), PUB011(bit2 excess combustion), PUB012(bit1 valve),
        PUB013(reset conditions), PUB014(bit2 only in overpressure), PUB015(continuous 3-scan)
*)
(* CONTRACT_RULES [] *)

tmpRisingReset := resetBtn AND NOT prevResetBtn;

tmpOverpressureValid := runRequest AND pressureValid AND (pressure >= 4500.0);

tmpStuckCond := tmpOverpressureValid AND (outletCmd >= 50) AND (outletFeedback <= 10);

tmpRisingPrevCond := prevRunRequest AND prevPressureValid AND (prevPressure >= 4500.0) AND (prevOutletCmd >= 50) AND (prevOutletFeedback <= 10);

tmpTwoAgoPrevCond := prevLatchedCauseMask; // placeholder, will use stored 2-ago state
tmpCurrentMask := 0;

IF NOT runRequest THEN
    tmpCurrentMask := 0;
    stuckValveConsecutiveCount := 0;
ELSIF NOT pressureValid THEN
    tmpCurrentMask := 1;
    stuckValveConsecutiveCount := 0;
ELSE
    IF tmpOverpressureValid THEN
        IF tmpStuckCond THEN
            IF tmpRisingPrevCond THEN
                stuckValveConsecutiveCount := 2;
            ELSE
                stuckValveConsecutiveCount := stuckValveConsecutiveCount + 1;
                IF stuckValveConsecutiveCount < 3 THEN
                    stuckValveConsecutiveCount := 3;
                END_IF;
            END_IF;
        ELSE
            stuckValveConsecutiveCount := 0;
        END_IF;

        IF stuckValveConsecutiveCount >= 3 THEN
            tmpCurrentMask := tmpCurrentMask OR 2;
        END_IF;

        IF (fuelFlow >= 4.0) AND (steamFlow <= 10.0) THEN
            tmpCurrentMask := tmpCurrentMask OR 4;
        END_IF;

        IF tmpCurrentMask = 0 THEN
            tmpCurrentMask := 8;
        END_IF;
    ELSE
        stuckValveConsecutiveCount := 0;
        tmpCurrentMask := 0;
    END_IF;
END_IF;

currentCauseMask := tmpCurrentMask;

IF tmpRisingReset AND NOT runRequest AND pressureValid AND (pressure <= 4200.0) THEN
    tripLatched := FALSE;
    latchedCauseMask := 0;
ELSIF runRequest AND (NOT pressureValid OR (pressure >= 4500.0)) THEN
    tripLatched := TRUE;
    latchedCauseMask := latchedCauseMask OR currentCauseMask;
ELSIF tripLatched THEN
    latchedCauseMask := latchedCauseMask OR currentCauseMask;
ELSE
    tripLatched := FALSE;
    latchedCauseMask := 0;
END_IF;

fuelPermit := runRequest AND NOT tripLatched;

diagnosticActive := (currentCauseMask <> 0);

prevResetBtn := resetBtn;
prevRunRequest := runRequest;
prevPressureValid := pressureValid;
prevPressure := pressure;
prevFuelFlow := fuelFlow;
prevSteamFlow := steamFlow;
prevOutletCmd := outletCmd;
prevOutletFeedback := outletFeedback;
prevTripLatched := tripLatched;
prevCurrentCauseMask := currentCauseMask;
prevLatchedCauseMask := latchedCauseMask;

END_FUNCTION_BLOCK
